   STAT29[4, 7].STAT30 := 0.000000e+000;
   STAT29[4, 7].STAT31 := 0.000000e+000;
   STAT29[4, 7].STAT32 := 0.000000e+000;
   STAT29[4, 8].STAT30 := 0.000000e+000;
   STAT29[4, 8].STAT31 := 0.000000e+000;
   STAT29[4, 8].STAT32 := 0.000000e+000;
   STAT29[4, 9].STAT30 := 0.000000e+000;
   STAT29[4, 9].STAT31 := 0.000000e+000;
   STAT29[4, 9].STAT32 := 0.000000e+000;
   STAT29[4, 10].STAT30 := 0.000000e+000;
   STAT29[4, 10].STAT31 := 0.000000e+000;
   STAT29[4, 10].STAT32 := 0.000000e+000;
   STAT29[5, 1].STAT30 := 0.000000e+000;
   STAT29[5, 1].STAT31 := 0.000000e+000;
   STAT29[5, 1].STAT32 := 0.000000e+000;
   STAT29[5, 2].STAT30 := 0.000000e+000;
   STAT29[5, 2].STAT31 := 0.000000e+000;
   STAT29[5, 2].STAT32 := 0.000000e+000;
   STAT29[5, 3].STAT30 := 0.000000e+000;
   STAT29[5, 3].STAT31 := 0.000000e+000;
   STAT29[5, 3].STAT32 := 0.000000e+000;
   STAT29[5, 4].STAT30 := 0.000000e+000;
   STAT29[5, 4].STAT31 := 0.000000e+000;
   STAT29[5, 4].STAT32 := 0.000000e+000;
   STAT29[5, 5].STAT30 := 0.000000e+000;
   STAT29[5, 5].STAT31 := 0.000000e+000;
   STAT29[5, 5].STAT32 := 0.000000e+000;
   STAT29[5, 6].STAT30 := 0.000000e+000;
   STAT29[5, 6].STAT31 := 0.000000e+000;
   STAT29[5, 6].STAT32 := 0.000000e+000;
   STAT29[5, 7].STAT30 := 0.000000e+000;
   STAT29[5, 7].STAT31 := 0.000000e+000;
   STAT29[5, 7].STAT32 := 0.000000e+000;
   STAT29[5, 8].STAT30 := 0.000000e+000;
   STAT29[5, 8].STAT31 := 0.000000e+000;
   STAT29[5, 8].STAT32 := 0.000000e+000;
   STAT29[5, 9].STAT30 := 0.000000e+000;
   STAT29[5, 9].STAT31 := 0.000000e+000;
   STAT29[5, 9].STAT32 := 0.000000e+000;
   STAT29[5, 10].STAT30 := 0.000000e+000;
   STAT29[5, 10].STAT31 := 0.000000e+000;
   STAT29[5, 10].STAT32 := 0.000000e+000;
   STAT29[6, 1].STAT30 := 0.000000e+000;
   STAT29[6, 1].STAT31 := 0.000000e+000;
   STAT29[6, 1].STAT32 := 0.000000e+000;
   STAT29[6, 2].STAT30 := 0.000000e+000;
   STAT29[6, 2].STAT31 := 0.000000e+000;
   STAT29[6, 2].STAT32 := 0.000000e+000;
   STAT29[6, 3].STAT30 := 0.000000e+000;
   STAT29[6, 3].STAT31 := 0.000000e+000;
   STAT29[6, 3].STAT32 := 0.000000e+000;
   STAT29[6, 4].STAT30 := 0.000000e+000;
   STAT29[6, 4].STAT31 := 0.000000e+000;
   STAT29[6, 4].STAT32 := 0.000000e+000;
   STAT29[6, 5].STAT30 := 0.000000e+000;
   STAT29[6, 5].STAT31 := 0.000000e+000;
   STAT29[6, 5].STAT32 := 0.000000e+000;
   STAT29[6, 6].STAT30 := 0.000000e+000;
   STAT29[6, 6].STAT31 := 0.000000e+000;
   STAT29[6, 6].STAT32 := 0.000000e+000;
   STAT29[6, 7].STAT30 := 0.000000e+000;
   STAT29[6, 7].STAT31 := 0.000000e+000;
   STAT29[6, 7].STAT32 := 0.000000e+000;
   STAT29[6, 8].STAT30 := 0.000000e+000;
   STAT29[6, 8].STAT31 := 0.000000e+000;
   STAT29[6, 8].STAT32 := 0.000000e+000;
   STAT29[6, 9].STAT30 := 0.000000e+000;
   STAT29[6, 9].STAT31 := 0.000000e+000;
   STAT29[6, 9].STAT32 := 0.000000e+000;
   STAT29[6, 10].STAT30 := 0.000000e+000;
   STAT29[6, 10].STAT31 := 0.000000e+000;
   STAT29[6, 10].STAT32 := 0.000000e+000;
   STAT29[7, 1].STAT30 := 0.000000e+000;
   STAT29[7, 1].STAT31 := 0.000000e+000;
   STAT29[7, 1].STAT32 := 0.000000e+000;
   STAT29[7, 2].STAT30 := 0.000000e+000;
   STAT29[7, 2].STAT31 := 0.000000e+000;
   STAT29[7, 2].STAT32 := 0.000000e+000;
   STAT29[7, 3].STAT30 := 0.000000e+000;
   STAT29[7, 3].STAT31 := 0.000000e+000;
   STAT29[7, 3].STAT32 := 0.000000e+000;
   STAT29[7, 4].STAT30 := 0.000000e+000;
   STAT29[7, 4].STAT31 := 0.000000e+000;
   STAT29[7, 4].STAT32 := 0.000000e+000;
   STAT29[7, 5].STAT30 := 0.000000e+000;
   STAT29[7, 5].STAT31 := 0.000000e+000;
   STAT29[7, 5].STAT32 := 0.000000e+000;
   STAT29[7, 6].STAT30 := 0.000000e+000;
   STAT29[7, 6].STAT31 := 0.000000e+000;
   STAT29[7, 6].STAT32 := 0.000000e+000;
   STAT29[7, 7].STAT30 := 0.000000e+000;
   STAT29[7, 7].STAT31 := 0.000000e+000;
   STAT29[7, 7].STAT32 := 0.000000e+000;
   STAT29[7, 8].STAT30 := 0.000000e+000;
   STAT29[7, 8].STAT31 := 0.000000e+000;
   STAT29[7, 8].STAT32 := 0.000000e+000;
   STAT29[7, 9].STAT30 := 0.000000e+000;
   STAT29[7, 9].STAT31 := 0.000000e+000;
   STAT29[7, 9].STAT32 := 0.000000e+000;
   STAT29[7, 10].STAT30 := 0.000000e+000;
   STAT29[7, 10].STAT31 := 0.000000e+000;
   STAT29[7, 10].STAT32 := 0.000000e+000;
   STAT29[8, 1].STAT30 := 0.000000e+000;
   STAT29[8, 1].STAT31 := 0.000000e+000;
   STAT29[8, 1].STAT32 := 0.000000e+000;
   STAT29[8, 2].STAT30 := 0.000000e+000;
   STAT29[8, 2].STAT31 := 0.000000e+000;
   STAT29[8, 2].STAT32 := 0.000000e+000;
   STAT29[8, 3].STAT30 := 0.000000e+000;
   STAT29[8, 3].STAT31 := 0.000000e+000;
   STAT29[8, 3].STAT32 := 0.000000e+000;
   STAT29[8, 4].STAT30 := 0.000000e+000;
   STAT29[8, 4].STAT31 := 0.000000e+000;
   STAT29[8, 4].STAT32 := 0.000000e+000;
   STAT29[8, 5].STAT30 := 0.000000e+000;
   STAT29[8, 5].STAT31 := 0.000000e+000;
   STAT29[8, 5].STAT32 := 0.000000e+000;
   STAT29[8, 6].STAT30 := 0.000000e+000;
   STAT29[8, 6].STAT31 := 0.000000e+000;
   STAT29[8, 6].STAT32 := 0.000000e+000;
   STAT29[8, 7].STAT30 := 0.000000e+000;
   STAT29[8, 7].STAT31 := 0.000000e+000;
   STAT29[8, 7].STAT32 := 0.000000e+000;
   STAT29[8, 8].STAT30 := 0.000000e+000;
   STAT29[8, 8].STAT31 := 0.000000e+000;
   STAT29[8, 8].STAT32 := 0.000000e+000;
   STAT29[8, 9].STAT30 := 0.000000e+000;
   STAT29[8, 9].STAT31 := 0.000000e+000;
   STAT29[8, 9].STAT32 := 0.000000e+000;
   STAT29[8, 10].STAT30 := 0.000000e+000;
   STAT29[8, 10].STAT31 := 0.000000e+000;
   STAT29[8, 10].STAT32 := 0.000000e+000;
   STAT29[9, 1].STAT30 := 0.000000e+000;
   STAT29[9, 1].STAT31 := 0.000000e+000;
   STAT29[9, 1].STAT32 := 0.000000e+000;
   STAT29[9, 2].STAT30 := 0.000000e+000;
   STAT29[9, 2].STAT31 := 0.000000e+000;
   STAT29[9, 2].STAT32 := 0.000000e+000;
   STAT29[9, 3].STAT30 := 0.000000e+000;
   STAT29[9, 3].STAT31 := 0.000000e+000;
   STAT29[9, 3].STAT32 := 0.000000e+000;
   STAT29[9, 4].STAT30 := 0.000000e+000;
   STAT29[9, 4].STAT31 := 0.000000e+000;
   STAT29[9, 4].STAT32 := 0.000000e+000;
   STAT29[9, 5].STAT30 := 0.000000e+000;
   STAT29[9, 5].STAT31 := 0.000000e+000;
   STAT29[9, 5].STAT32 := 0.000000e+000;
   STAT29[9, 6].STAT30 := 0.000000e+000;
   STAT29[9, 6].STAT31 := 0.000000e+000;
   STAT29[9, 6].STAT32 := 0.000000e+000;
   STAT29[9, 7].STAT30 := 0.000000e+000;
   STAT29[9, 7].STAT31 := 0.000000e+000;
   STAT29[9, 7].STAT32 := 0.000000e+000;
   STAT29[9, 8].STAT30 := 0.000000e+000;
   STAT29[9, 8].STAT31 := 0.000000e+000;
   STAT29[9, 8].STAT32 := 0.000000e+000;
   STAT29[9, 9].STAT30 := 0.000000e+000;
   STAT29[9, 9].STAT31 := 0.000000e+000;
   STAT29[9, 9].STAT32 := 0.000000e+000;
   STAT29[9, 10].STAT30 := 0.000000e+000;
   STAT29[9, 10].STAT31 := 0.000000e+000;
   STAT29[9, 10].STAT32 := 0.000000e+000;
   STAT29[10, 1].STAT30 := 0.000000e+000;
   STAT29[10, 1].STAT31 := 0.000000e+000;
   STAT29[10, 1].STAT32 := 0.000000e+000;
   STAT29[10, 2].STAT30 := 0.000000e+000;
   STAT29[10, 2].STAT31 := 0.000000e+000;
   STAT29[10, 2].STAT32 := 0.000000e+000;
   STAT29[10, 3].STAT30 := 0.000000e+000;
   STAT29[10, 3].STAT31 := 0.000000e+000;
   STAT29[10, 3].STAT32 := 0.000000e+000;
   STAT29[10, 4].STAT30 := 0.000000e+000;
   STAT29[10, 4].STAT31 := 0.000000e+000;
   STAT29[10, 4].STAT32 := 0.000000e+000;
   STAT29[10, 5].STAT30 := 0.000000e+000;
   STAT29[10, 5].STAT31 := 0.000000e+000;
   STAT29[10, 5].STAT32 := 0.000000e+000;
   STAT29[10, 6].STAT30 := 0.000000e+000;
   STAT29[10, 6].STAT31 := 0.000000e+000;
   STAT29[10, 6].STAT32 := 0.000000e+000;
   STAT29[10, 7].STAT30 := 0.000000e+000;
   STAT29[10, 7].STAT31 := 0.000000e+000;
   STAT29[10, 7].STAT32 := 0.000000e+000;
   STAT29[10, 8].STAT30 := 0.000000e+000;
   STAT29[10, 8].STAT31 := 0.000000e+000;
   STAT29[10, 8].STAT32 := 0.000000e+000;
   STAT29[10, 9].STAT30 := 0.000000e+000;
   STAT29[10, 9].STAT31 := 0.000000e+000;
   STAT29[10, 9].STAT32 := 0.000000e+000;
   STAT29[10, 10].STAT30 := 0.000000e+000;
   STAT29[10, 10].STAT31 := 0.000000e+000;
   STAT29[10, 10].STAT32 := 0.000000e+000;
   STAT33[1, 1, 1] := 0.000000e+000;
   STAT33[1, 1, 2] := 0.000000e+000;
   STAT33[1, 1, 3] := 0.000000e+000;
   STAT33[1, 1, 4] := 0.000000e+000;
   STAT33[1, 1, 5] := 0.000000e+000;
   STAT33[1, 1, 6] := 0.000000e+000;
   STAT33[1, 1, 7] := 0.000000e+000;
   STAT33[1, 1, 8] := 0.000000e+000;
   STAT33[1, 1, 9] := 0.000000e+000;
   STAT33[1, 1, 10] := 0.000000e+000;
   STAT33[1, 2, 1] := 0.000000e+000;
   STAT33[1, 2, 2] := 0.000000e+000;
   STAT33[1, 2, 3] := 0.000000e+000;
   STAT33[1, 2, 4] := 0.000000e+000;
   STAT33[1, 2, 5] := 0.000000e+000;
   STAT33[1, 2, 6] := 0.000000e+000;
   STAT33[1, 2, 7] := 0.000000e+000;
   STAT33[1, 2, 8] := 0.000000e+000;
   STAT33[1, 2, 9] := 0.000000e+000;
   STAT33[1, 2, 10] := 0.000000e+000;
   STAT33[1, 3, 1] := 0.000000e+000;
   STAT33[1, 3, 2] := 0.000000e+000;
   STAT33[1, 3, 3] := 0.000000e+000;
   STAT33[1, 3, 4] := 0.000000e+000;
   STAT33[1, 3, 5] := 0.000000e+000;
   STAT33[1, 3, 6] := 0.000000e+000;
   STAT33[1, 3, 7] := 0.000000e+000;
   STAT33[1, 3, 8] := 0.000000e+000;
   STAT33[1, 3, 9] := 0.000000e+000;
   STAT33[1, 3, 10] := 0.000000e+000;
   STAT33[1, 4, 1] := 0.000000e+000;
   STAT33[1, 4, 2] := 0.000000e+000;
   STAT33[1, 4, 3] := 0.000000e+000;
   STAT33[1, 4, 4] := 0.000000e+000;
   STAT33[1, 4, 5] := 0.000000e+000;
   STAT33[1, 4, 6] := 0.000000e+000;
   STAT33[1, 4, 7] := 0.000000e+000;
   STAT33[1, 4, 8] := 0.000000e+000;
   STAT33[1, 4, 9] := 0.000000e+000;
   STAT33[1, 4, 10] := 0.000000e+000;
   STAT33[1, 5, 1] := 0.000000e+000;
   STAT33[1, 5, 2] := 0.000000e+000;
   STAT33[1, 5, 3] := 0.000000e+000;
   STAT33[1, 5, 4] := 0.000000e+000;
   STAT33[1, 5, 5] := 0.000000e+000;
   STAT33[1, 5, 6] := 0.000000e+000;
   STAT33[1, 5, 7] := 0.000000e+000;
   STAT33[1, 5, 8] := 0.000000e+000;
   STAT33[1, 5, 9] := 0.000000e+000;
   STAT33[1, 5, 10] := 0.000000e+000;
   STAT33[1, 6, 1] := 0.000000e+000;
   STAT33[1, 6, 2] := 0.000000e+000;
   STAT33[1, 6, 3] := 0.000000e+000;
   STAT33[1, 6, 4] := 0.000000e+000;
   STAT33[1, 6, 5] := 0.000000e+000;
   STAT33[1, 6, 6] := 0.000000e+000;
   STAT33[1, 6, 7] := 0.000000e+000;
   STAT33[1, 6, 8] := 0.000000e+000;
   STAT33[1, 6, 9] := 0.000000e+000;
   STAT33[1, 6, 10] := 0.000000e+000;
   STAT33[1, 7, 1] := 0.000000e+000;
   STAT33[1, 7, 2] := 0.000000e+000;
   STAT33[1, 7, 3] := 0.000000e+000;
   STAT33[1, 7, 4] := 0.000000e+000;
   STAT33[1, 7, 5] := 0.000000e+000;
   STAT33[1, 7, 6] := 0.000000e+000;
   STAT33[1, 7, 7] := 0.000000e+000;
   STAT33[1, 7, 8] := 0.000000e+000;
   STAT33[1, 7, 9] := 0.000000e+000;
   STAT33[1, 7, 10] := 0.000000e+000;
   STAT33[1, 8, 1] := 0.000000e+000;
   STAT33[1, 8, 2] := 0.000000e+000;
   STAT33[1, 8, 3] := 0.000000e+000;
   STAT33[1, 8, 4] := 0.000000e+000;
   STAT33[1, 8, 5] := 0.000000e+000;
   STAT33[1, 8, 6] := 0.000000e+000;
   STAT33[1, 8, 7] := 0.000000e+000;
   STAT33[1, 8, 8] := 0.000000e+000;
   STAT33[1, 8, 9] := 0.000000e+000;
   STAT33[1, 8, 10] := 0.000000e+000;
   STAT33[1, 9, 1] := 0.000000e+000;
   STAT33[1, 9, 2] := 0.000000e+000;
   STAT33[1, 9, 3] := 0.000000e+000;
   STAT33[1, 9, 4] := 0.000000e+000;
   STAT33[1, 9, 5] := 0.000000e+000;
   STAT33[1, 9, 6] := 0.000000e+000;
   STAT33[1, 9, 7] := 0.000000e+000;
   STAT33[1, 9, 8] := 0.000000e+000;
   STAT33[1, 9, 9] := 0.000000e+000;
   STAT33[1, 9, 10] := 0.000000e+000;
   STAT33[1, 10, 1] := 0.000000e+000;
   STAT33[1, 10, 2] := 0.000000e+000;
   STAT33[1, 10, 3] := 0.000000e+000;
   STAT33[1, 10, 4] := 0.000000e+000;
   STAT33[1, 10, 5] := 0.000000e+000;
   STAT33[1, 10, 6] := 0.000000e+000;
   STAT33[1, 10, 7] := 0.000000e+000;
   STAT33[1, 10, 8] := 0.000000e+000;
   STAT33[1, 10, 9] := 0.000000e+000;
   STAT33[1, 10, 10] := 0.000000e+000;
   STAT33[2, 1, 1] := 0.000000e+000;
   STAT33[2, 1, 2] := 0.000000e+000;
   STAT33[2, 1, 3] := 0.000000e+000;
   STAT33[2, 1, 4] := 0.000000e+000;
   STAT33[2, 1, 5] := 0.000000e+000;
   STAT33[2, 1, 6] := 0.000000e+000;
   STAT33[2, 1, 7] := 0.000000e+000;
   STAT33[2, 1, 8] := 0.000000e+000;
   STAT33[2, 1, 9] := 0.000000e+000;
   STAT33[2, 1, 10] := 0.000000e+000;
   STAT33[2, 2, 1] := 0.000000e+000;
   STAT33[2, 2, 2] := 0.000000e+000;
   STAT33[2, 2, 3] := 0.000000e+000;
   STAT33[2, 2, 4] := 0.000000e+000;
   STAT33[2, 2, 5] := 0.000000e+000;
   STAT33[2, 2, 6] := 0.000000e+000;
   STAT33[2, 2, 7] := 0.000000e+000;
   STAT33[2, 2, 8] := 0.000000e+000;
   STAT33[2, 2, 9] := 0.000000e+000;
   STAT33[2, 2, 10] := 0.000000e+000;
   STAT33[2, 3, 1] := 0.000000e+000;
   STAT33[2, 3, 2] := 0.000000e+000;
   STAT33[2, 3, 3] := 0.000000e+000;
   STAT33[2, 3, 4] := 0.000000e+000;
   STAT33[2, 3, 5] := 0.000000e+000;
   STAT33[2, 3, 6] := 0.000000e+000;
   STAT33[2, 3, 7] := 0.000000e+000;
   STAT33[2, 3, 8] := 0.000000e+000;
   STAT33[2, 3, 9] := 0.000000e+000;
   STAT33[2, 3, 10] := 0.000000e+000;
   STAT33[2, 4, 1] := 0.000000e+000;
   STAT33[2, 4, 2] := 0.000000e+000;
   STAT33[2, 4, 3] := 0.000000e+000;
   STAT33[2, 4, 4] := 0.000000e+000;
   STAT33[2, 4, 5] := 0.000000e+000;
   STAT33[2, 4, 6] := 0.000000e+000;
   STAT33[2, 4, 7] := 0.000000e+000;
   STAT33[2, 4, 8] := 0.000000e+000;
   STAT33[2, 4, 9] := 0.000000e+000;
   STAT33[2, 4, 10] := 0.000000e+000;
   STAT33[2, 5, 1] := 0.000000e+000;
   STAT33[2, 5, 2] := 0.000000e+000;
   STAT33[2, 5, 3] := 0.000000e+000;
   STAT33[2, 5, 4] := 0.000000e+000;
   STAT33[2, 5, 5] := 0.000000e+000;
   STAT33[2, 5, 6] := 0.000000e+000;
   STAT33[2, 5, 7] := 0.000000e+000;
   STAT33[2, 5, 8] := 0.000000e+000;
   STAT33[2, 5, 9] := 0.000000e+000;
   STAT33[2, 5, 10] := 0.000000e+000;
   STAT33[2, 6, 1] := 0.000000e+000;
   STAT33[2, 6, 2] := 0.000000e+000;
   STAT33[2, 6, 3] := 0.000000e+000;
   STAT33[2, 6, 4] := 0.000000e+000;
   STAT33[2, 6, 5] := 0.000000e+000;
   STAT33[2, 6, 6] := 0.000000e+000;
   STAT33[2, 6, 7] := 0.000000e+000;
   STAT33[2, 6, 8] := 0.000000e+000;
   STAT33[2, 6, 9] := 0.000000e+000;
   STAT33[2, 6, 10] := 0.000000e+000;
   STAT33[2, 7, 1] := 0.000000e+000;
   STAT33[2, 7, 2] := 0.000000e+000;
   STAT33[2, 7, 3] := 0.000000e+000;
   STAT33[2, 7, 4] := 0.000000e+000;
   STAT33[2, 7, 5] := 0.000000e+000;
   STAT33[2, 7, 6] := 0.000000e+000;
   STAT33[2, 7, 7] := 0.000000e+000;
   STAT33[2, 7, 8] := 0.000000e+000;
   STAT33[2, 7, 9] := 0.000000e+000;
   STAT33[2, 7, 10] := 0.000000e+000;
   STAT33[2, 8, 1] := 0.000000e+000;
   STAT33[2, 8, 2] := 0.000000e+000;
   STAT33[2, 8, 3] := 0.000000e+000;
   STAT33[2, 8, 4] := 0.000000e+000;
   STAT33[2, 8, 5] := 0.000000e+000;
   STAT33[2, 8, 6] := 0.000000e+000;
   STAT33[2, 8, 7] := 0.000000e+000;
   STAT33[2, 8, 8] := 0.000000e+000;
   STAT33[2, 8, 9] := 0.000000e+000;
   STAT33[2, 8, 10] := 0.000000e+000;
   STAT33[2, 9, 1] := 0.000000e+000;
   STAT33[2, 9, 2] := 0.000000e+000;
   STAT33[2, 9, 3] := 0.000000e+000;
   STAT33[2, 9, 4] := 0.000000e+000;
   STAT33[2, 9, 5] := 0.000000e+000;
   STAT33[2, 9, 6] := 0.000000e+000;
   STAT33[2, 9, 7] := 0.000000e+000;
   STAT33[2, 9, 8] := 0.000000e+000;
   STAT33[2, 9, 9] := 0.000000e+000;
   STAT33[2, 9, 10] := 0.000000e+000;
   STAT33[2, 10, 1] := 0.000000e+000;
   STAT33[2, 10, 2] := 0.000000e+000;
   STAT33[2, 10, 3] := 0.000000e+000;
   STAT33[2, 10, 4] := 0.000000e+000;
   STAT33[2, 10, 5] := 0.000000e+000;
   STAT33[2, 10, 6] := 0.000000e+000;
   STAT33[2, 10, 7] := 0.000000e+000;
   STAT33[2, 10, 8] := 0.000000e+000;
   STAT33[2, 10, 9] := 0.000000e+000;
   STAT33[2, 10, 10] := 0.000000e+000;
   STAT33[3, 1, 1] := 0.000000e+000;
   STAT33[3, 1, 2] := 0.000000e+000;
   STAT33[3, 1, 3] := 0.000000e+000;
   STAT33[3, 1, 4] := 0.000000e+000;
   STAT33[3, 1, 5] := 0.000000e+000;
   STAT33[3, 1, 6] := 0.000000e+000;
   STAT33[3, 1, 7] := 0.000000e+000;
   STAT33[3, 1, 8] := 0.000000e+000;
   STAT33[3, 1, 9] := 0.000000e+000;
   STAT33[3, 1, 10] := 0.000000e+000;
   STAT33[3, 2, 1] := 0.000000e+000;
   STAT33[3, 2, 2] := 0.000000e+000;
   STAT33[3, 2, 3] := 0.000000e+000;
   STAT33[3, 2, 4] := 0.000000e+000;
   STAT33[3, 2, 5] := 0.000000e+000;
   STAT33[3, 2, 6] := 0.000000e+000;
   STAT33[3, 2, 7] := 0.000000e+000;
   STAT33[3, 2, 8] := 0.000000e+000;
   STAT33[3, 2, 9] := 0.000000e+000;
   STAT33[3, 2, 10] := 0.000000e+000;
   STAT33[3, 3, 1] := 0.000000e+000;
   STAT33[3, 3, 2] := 0.000000e+000;
   STAT33[3, 3, 3] := 0.000000e+000;
   STAT33[3, 3, 4] := 0.000000e+000;
   STAT33[3, 3, 5] := 0.000000e+000;
   STAT33[3, 3, 6] := 0.000000e+000;
   STAT33[3, 3, 7] := 0.000000e+000;
   STAT33[3, 3, 8] := 0.000000e+000;
   STAT33[3, 3, 9] := 0.000000e+000;
   STAT33[3, 3, 10] := 0.000000e+000;
   STAT33[3, 4, 1] := 0.000000e+000;
   STAT33[3, 4, 2] := 0.000000e+000;
   STAT33[3, 4, 3] := 0.000000e+000;
   STAT33[3, 4, 4] := 0.000000e+000;
   STAT33[3, 4, 5] := 0.000000e+000;
   STAT33[3, 4, 6] := 0.000000e+000;
   STAT33[3, 4, 7] := 0.000000e+000;
   STAT33[3, 4, 8] := 0.000000e+000;
   STAT33[3, 4, 9] := 0.000000e+000;
   STAT33[3, 4, 10] := 0.000000e+000;
   STAT33[3, 5, 1] := 0.000000e+000;
   STAT33[3, 5, 2] := 0.000000e+000;
   STAT33[3, 5, 3] := 0.000000e+000;
   STAT33[3, 5, 4] := 0.000000e+000;
   STAT33[3, 5, 5] := 0.000000e+000;
   STAT33[3, 5, 6] := 0.000000e+000;
   STAT33[3, 5, 7] := 0.000000e+000;
   STAT33[3, 5, 8] := 0.000000e+000;
   STAT33[3, 5, 9] := 0.000000e+000;
   STAT33[3, 5, 10] := 0.000000e+000;
   STAT33[3, 6, 1] := 0.000000e+000;
   STAT33[3, 6, 2] := 0.000000e+000;
   STAT33[3, 6, 3] := 0.000000e+000;
   STAT33[3, 6, 4] := 0.000000e+000;
   STAT33[3, 6, 5] := 0.000000e+000;
   STAT33[3, 6, 6] := 0.000000e+000;
   STAT33[3, 6, 7] := 0.000000e+000;
   STAT33[3, 6, 8] := 0.000000e+000;
   STAT33[3, 6, 9] := 0.000000e+000;
   STAT33[3, 6, 10] := 0.000000e+000;
   STAT33[3, 7, 1] := 0.000000e+000;
   STAT33[3, 7, 2] := 0.000000e+000;
   STAT33[3, 7, 3] := 0.000000e+000;
   STAT33[3, 7, 4] := 0.000000e+000;
   STAT33[3, 7, 5] := 0.000000e+000;
   STAT33[3, 7, 6] := 0.000000e+000;
   STAT33[3, 7, 7] := 0.000000e+000;
   STAT33[3, 7, 8] := 0.000000e+000;
   STAT33[3, 7, 9] := 0.000000e+000;
   STAT33[3, 7, 10] := 0.000000e+000;
   STAT33[3, 8, 1] := 0.000000e+000;
   STAT33[3, 8, 2] := 0.000000e+000;
   STAT33[3, 8, 3] := 0.000000e+000;
   STAT33[3, 8, 4] := 0.000000e+000;
   STAT33[3, 8, 5] := 0.000000e+000;
   STAT33[3, 8, 6] := 0.000000e+000;
   STAT33[3, 8, 7] := 0.000000e+000;
   STAT33[3, 8, 8] := 0.000000e+000;
   STAT33[3, 8, 9] := 0.000000e+000;
   STAT33[3, 8, 10] := 0.000000e+000;
   STAT33[3, 9, 1] := 0.000000e+000;
   STAT33[3, 9, 2] := 0.000000e+000;
   STAT33[3, 9, 3] := 0.000000e+000;
   STAT33[3, 9, 4] := 0.000000e+000;
   STAT33[3, 9, 5] := 0.000000e+000;
   STAT33[3, 9, 6] := 0.000000e+000;
   STAT33[3, 9, 7] := 0.000000e+000;
   STAT33[3, 9, 8] := 0.000000e+000;
   STAT33[3, 9, 9] := 0.000000e+000;
   STAT33[3, 9, 10] := 0.000000e+000;
   STAT33[3, 10, 1] := 0.000000e+000;
   STAT33[3, 10, 2] := 0.000000e+000;
   STAT33[3, 10, 3] := 0.000000e+000;
   STAT33[3, 10, 4] := 0.000000e+000;
   STAT33[3, 10, 5] := 0.000000e+000;
   STAT33[3, 10, 6] := 0.000000e+000;
   STAT33[3, 10, 7] := 0.000000e+000;
   STAT33[3, 10, 8] := 0.000000e+000;
   STAT33[3, 10, 9] := 0.000000e+000;
   STAT33[3, 10, 10] := 0.000000e+000;
   STAT33[4, 1, 1] := 0.000000e+000;
   STAT33[4, 1, 2] := 0.000000e+000;
   STAT33[4, 1, 3] := 0.000000e+000;
   STAT33[4, 1, 4] := 0.000000e+000;
   STAT33[4, 1, 5] := 0.000000e+000;
   STAT33[4, 1, 6] := 0.000000e+000;
   STAT33[4, 1, 7] := 0.000000e+000;
   STAT33[4, 1, 8] := 0.000000e+000;
   STAT33[4, 1, 9] := 0.000000e+000;
   STAT33[4, 1, 10] := 0.000000e+000;
   STAT33[4, 2, 1] := 0.000000e+000;
   STAT33[4, 2, 2] := 0.000000e+000;
   STAT33[4, 2, 3] := 0.000000e+000;
   STAT33[4, 2, 4] := 0.000000e+000;
   STAT33[4, 2, 5] := 0.000000e+000;
   STAT33[4, 2, 6] := 0.000000e+000;
   STAT33[4, 2, 7] := 0.000000e+000;
   STAT33[4, 2, 8] := 0.000000e+000;
   STAT33[4, 2, 9] := 0.000000e+000;
   STAT33[4, 2, 10] := 0.000000e+000;
   STAT33[4, 3, 1] := 0.000000e+000;
   STAT33[4, 3, 2] := 0.000000e+000;
   STAT33[4, 3, 3] := 0.000000e+000;
   STAT33[4, 3, 4] := 0.000000e+000;
   STAT33[4, 3, 5] := 0.000000e+000;
   STAT33[4, 3, 6] := 0.000000e+000;
   STAT33[4, 3, 7] := 0.000000e+000;
   STAT33[4, 3, 8] := 0.000000e+000;
   STAT33[4, 3, 9] := 0.000000e+000;
   STAT33[4, 3, 10] := 0.000000e+000;
   STAT33[4, 4, 1] := 0.000000e+000;
   STAT33[4, 4, 2] := 0.000000e+000;
   STAT33[4, 4, 3] := 0.000000e+000;
   STAT33[4, 4, 4] := 0.000000e+000;
   STAT33[4, 4, 5] := 0.000000e+000;
   STAT33[4, 4, 6] := 0.000000e+000;
   STAT33[4, 4, 7] := 0.000000e+000;
   STAT33[4, 4, 8] := 0.000000e+000;
   STAT33[4, 4, 9] := 0.000000e+000;
   STAT33[4, 4, 10] := 0.000000e+000;
   STAT33[4, 5, 1] := 0.000000e+000;
   STAT33[4, 5, 2] := 0.000000e+000;
   STAT33[4, 5, 3] := 0.000000e+000;
   STAT33[4, 5, 4] := 0.000000e+000;
   STAT33[4, 5, 5] := 0.000000e+000;
   STAT33[4, 5, 6] := 0.000000e+000;
   STAT33[4, 5, 7] := 0.000000e+000;
   STAT33[4, 5, 8] := 0.000000e+000;
   STAT33[4, 5, 9] := 0.000000e+000;
   STAT33[4, 5, 10] := 0.000000e+000;
   STAT33[4, 6, 1] := 0.000000e+000;
   STAT33[4, 6, 2] := 0.000000e+000;
   STAT33[4, 6, 3] := 0.000000e+000;
   STAT33[4, 6, 4] := 0.000000e+000;
   STAT33[4, 6, 5] := 0.000000e+000;
   STAT33[4, 6, 6] := 0.000000e+000;
   STAT33[4, 6, 7] := 0.000000e+000;
   STAT33[4, 6, 8] := 0.000000e+000;
   STAT33[4, 6, 9] := 0.000000e+000;
   STAT33[4, 6, 10] := 0.000000e+000;
   STAT33[4, 7, 1] := 0.000000e+000;
   STAT33[4, 7, 2] := 0.000000e+000;
   STAT33[4, 7, 3] := 0.000000e+000;
   STAT33[4, 7, 4] := 0.000000e+000;
   STAT33[4, 7, 5] := 0.000000e+000;
   STAT33[4, 7, 6] := 0.000000e+000;
   STAT33[4, 7, 7] := 0.000000e+000;
   STAT33[4, 7, 8] := 0.000000e+000;
   STAT33[4, 7, 9] := 0.000000e+000;
   STAT33[4, 7, 10] := 0.000000e+000;
   STAT33[4, 8, 1] := 0.000000e+000;
   STAT33[4, 8, 2] := 0.000000e+000;
   STAT33[4, 8, 3] := 0.000000e+000;
   STAT33[4, 8, 4] := 0.000000e+000;
   STAT33[4, 8, 5] := 0.000000e+000;
   STAT33[4, 8, 6] := 0.000000e+000;
   STAT33[4, 8, 7] := 0.000000e+000;
   STAT33[4, 8, 8] := 0.000000e+000;
   STAT33[4, 8, 9] := 0.000000e+000;
   STAT33[4, 8, 10] := 0.000000e+000;
   STAT33[4, 9, 1] := 0.000000e+000;
   STAT33[4, 9, 2] := 0.000000e+000;
   STAT33[4, 9, 3] := 0.000000e+000;
   STAT33[4, 9, 4] := 0.000000e+000;
   STAT33[4, 9, 5] := 0.000000e+000;
   STAT33[4, 9, 6] := 0.000000e+000;
   STAT33[4, 9, 7] := 0.000000e+000;
   STAT33[4, 9, 8] := 0.000000e+000;
   STAT33[4, 9, 9] := 0.000000e+000;
   STAT33[4, 9, 10] := 0.000000e+000;
   STAT33[4, 10, 1] := 0.000000e+000;
   STAT33[4, 10, 2] := 0.000000e+000;
   STAT33[4, 10, 3] := 0.000000e+000;
   STAT33[4, 10, 4] := 0.000000e+000;
   STAT33[4, 10, 5] := 0.000000e+000;
   STAT33[4, 10, 6] := 0.000000e+000;
   STAT33[4, 10, 7] := 0.000000e+000;
   STAT33[4, 10, 8] := 0.000000e+000;
   STAT33[4, 10, 9] := 0.000000e+000;
   STAT33[4, 10, 10] := 0.000000e+000;
   STAT33[5, 1, 1] := 0.000000e+000;
   STAT33[5, 1, 2] := 0.000000e+000;
   STAT33[5, 1, 3] := 0.000000e+000;
   STAT33[5, 1, 4] := 0.000000e+000;
   STAT33[5, 1, 5] := 0.000000e+000;
   STAT33[5, 1, 6] := 0.000000e+000;
   STAT33[5, 1, 7] := 0.000000e+000;
   STAT33[5, 1, 8] := 0.000000e+000;
   STAT33[5, 1, 9] := 0.000000e+000;
   STAT33[5, 1, 10] := 0.000000e+000;
   STAT33[5, 2, 1] := 0.000000e+000;
   STAT33[5, 2, 2] := 0.000000e+000;
   STAT33[5, 2, 3] := 0.000000e+000;
   STAT33[5, 2, 4] := 0.000000e+000;
   STAT33[5, 2, 5] := 0.000000e+000;
   STAT33[5, 2, 6] := 0.000000e+000;
   STAT33[5, 2, 7] := 0.000000e+000;
   STAT33[5, 2, 8] := 0.000000e+000;
   STAT33[5, 2, 9] := 0.000000e+000;
   STAT33[5, 2, 10] := 0.000000e+000;
   STAT33[5, 3, 1] := 0.000000e+000;
   STAT33[5, 3, 2] := 0.000000e+000;
   STAT33[5, 3, 3] := 0.000000e+000;
   STAT33[5, 3, 4] := 0.000000e+000;
   STAT33[5, 3, 5] := 0.000000e+000;
   STAT33[5, 3, 6] := 0.000000e+000;
   STAT33[5, 3, 7] := 0.000000e+000;
   STAT33[5, 3, 8] := 0.000000e+000;
   STAT33[5, 3, 9] := 0.000000e+000;
   STAT33[5, 3, 10] := 0.000000e+000;
   STAT33[5, 4, 1] := 0.000000e+000;
   STAT33[5, 4, 2] := 0.000000e+000;
   STAT33[5, 4, 3] := 0.000000e+000;
   STAT33[5, 4, 4] := 0.000000e+000;
   STAT33[5, 4, 5] := 0.000000e+000;
   STAT33[5, 4, 6] := 0.000000e+000;
   STAT33[5, 4, 7] := 0.000000e+000;
   STAT33[5, 4, 8] := 0.000000e+000;
   STAT33[5, 4, 9] := 0.000000e+000;
   STAT33[5, 4, 10] := 0.000000e+000;
   STAT33[5, 5, 1] := 0.000000e+000;
   STAT33[5, 5, 2] := 0.000000e+000;
   STAT33[5, 5, 3] := 0.000000e+000;
   STAT33[5, 5, 4] := 0.000000e+000;
   STAT33[5, 5, 5] := 0.000000e+000;
   STAT33[5, 5, 6] := 0.000000e+000;
   STAT33[5, 5, 7] := 0.000000e+000;
   STAT33[5, 5, 8] := 0.000000e+000;
   STAT33[5, 5, 9] := 0.000000e+000;
   STAT33[5, 5, 10] := 0.000000e+000;
   STAT33[5, 6, 1] := 0.000000e+000;
   STAT33[5, 6, 2] := 0.000000e+000;
   STAT33[5, 6, 3] := 0.000000e+000;
   STAT33[5, 6, 4] := 0.000000e+000;
   STAT33[5, 6, 5] := 0.000000e+000;
   STAT33[5, 6, 6] := 0.000000e+000;
   STAT33[5, 6, 7] := 0.000000e+000;
   STAT33[5, 6, 8] := 0.000000e+000;
   STAT33[5, 6, 9] := 0.000000e+000;
   STAT33[5, 6, 10] := 0.000000e+000;
   STAT33[5, 7, 1] := 0.000000e+000;
   STAT33[5, 7, 2] := 0.000000e+000;
   STAT33[5, 7, 3] := 0.000000e+000;
   STAT33[5, 7, 4] := 0.000000e+000;
   STAT33[5, 7, 5] := 0.000000e+000;
   STAT33[5, 7, 6] := 0.000000e+000;
   STAT33[5, 7, 7] := 0.000000e+000;
   STAT33[5, 7, 8] := 0.000000e+000;
   STAT33[5, 7, 9] := 0.000000e+000;
   STAT33[5, 7, 10] := 0.000000e+000;
   STAT33[5, 8, 1] := 0.000000e+000;
   STAT33[5, 8, 2] := 0.000000e+000;
   STAT33[5, 8, 3] := 0.000000e+000;
   STAT33[5, 8, 4] := 0.000000e+000;
   STAT33[5, 8, 5] := 0.000000e+000;
   STAT33[5, 8, 6] := 0.000000e+000;
   STAT33[5, 8, 7] := 0.000000e+000;
   STAT33[5, 8, 8] := 0.000000e+000;
   STAT33[5, 8, 9] := 0.000000e+000;
   STAT33[5, 8, 10] := 0.000000e+000;
   STAT33[5, 9, 1] := 0.000000e+000;
   STAT33[5, 9, 2] := 0.000000e+000;
   STAT33[5, 9, 3] := 0.000000e+000;
   STAT33[5, 9, 4] := 0.000000e+000;
   STAT33[5, 9, 5] := 0.000000e+000;
   STAT33[5, 9, 6] := 0.000000e+000;
   STAT33[5, 9, 7] := 0.000000e+000;
   STAT33[5, 9, 8] := 0.000000e+000;
   STAT33[5, 9, 9] := 0.000000e+000;
   STAT33[5, 9, 10] := 0.000000e+000;
   STAT33[5, 10, 1] := 0.000000e+000;
   STAT33[5, 10, 2] := 0.000000e+000;
   STAT33[5, 10, 3] := 0.000000e+000;
   STAT33[5, 10, 4] := 0.000000e+000;
   STAT33[5, 10, 5] := 0.000000e+000;
   STAT33[5, 10, 6] := 0.000000e+000;
   STAT33[5, 10, 7] := 0.000000e+000;
   STAT33[5, 10, 8] := 0.000000e+000;
   STAT33[5, 10, 9] := 0.000000e+000;
   STAT33[5, 10, 10] := 0.000000e+000;
   STAT33[6, 1, 1] := 0.000000e+000;
   STAT33[6, 1, 2] := 0.000000e+000;
   STAT33[6, 1, 3] := 0.000000e+000;
   STAT33[6, 1, 4] := 0.000000e+000;
   STAT33[6, 1, 5] := 0.000000e+000;
   STAT33[6, 1, 6] := 0.000000e+000;
   STAT33[6, 1, 7] := 0.000000e+000;
   STAT33[6, 1, 8] := 0.000000e+000;
   STAT33[6, 1, 9] := 0.000000e+000;
   STAT33[6, 1, 10] := 0.000000e+000;
   STAT33[6, 2, 1] := 0.000000e+000;
   STAT33[6, 2, 2] := 0.000000e+000;
   STAT33[6, 2, 3] := 0.000000e+000;
   STAT33[6, 2, 4] := 0.000000e+000;
   STAT33[6, 2, 5] := 0.000000e+000;
   STAT33[6, 2, 6] := 0.000000e+000;
   STAT33[6, 2, 7] := 0.000000e+000;
   STAT33[6, 2, 8] := 0.000000e+000;
   STAT33[6, 2, 9] := 0.000000e+000;
   STAT33[6, 2, 10] := 0.000000e+000;
   STAT33[6, 3, 1] := 0.000000e+000;
   STAT33[6, 3, 2] := 0.000000e+000;
   STAT33[6, 3, 3] := 0.000000e+000;
   STAT33[6, 3, 4] := 0.000000e+000;
   STAT33[6, 3, 5] := 0.000000e+000;
   STAT33[6, 3, 6] := 0.000000e+000;
   STAT33[6, 3, 7] := 0.000000e+000;
   STAT33[6, 3, 8] := 0.000000e+000;
   STAT33[6, 3, 9] := 0.000000e+000;
   STAT33[6, 3, 10] := 0.000000e+000;
   STAT33[6, 4, 1] := 0.000000e+000;
   STAT33[6, 4, 2] := 0.000000e+000;
   STAT33[6, 4, 3] := 0.000000e+000;
   STAT33[6, 4, 4] := 0.000000e+000;
   STAT33[6, 4, 5] := 0.000000e+000;
   STAT33[6, 4, 6] := 0.000000e+000;
   STAT33[6, 4, 7] := 0.000000e+000;
   STAT33[6, 4, 8] := 0.000000e+000;
   STAT33[6, 4, 9] := 0.000000e+000;
   STAT33[6, 4, 10] := 0.000000e+000;
   STAT33[6, 5, 1] := 0.000000e+000;
   STAT33[6, 5, 2] := 0.000000e+000;
   STAT33[6, 5, 3] := 0.000000e+000;
   STAT33[6, 5, 4] := 0.000000e+000;
   STAT33[6, 5, 5] := 0.000000e+000;
   STAT33[6, 5, 6] := 0.000000e+000;
   STAT33[6, 5, 7] := 0.000000e+000;
   STAT33[6, 5, 8] := 0.000000e+000;
   STAT33[6, 5, 9] := 0.000000e+000;
   STAT33[6, 5, 10] := 0.000000e+000;
   STAT33[6, 6, 1] := 0.000000e+000;
   STAT33[6, 6, 2] := 0.000000e+000;
   STAT33[6, 6, 3] := 0.000000e+000;
   STAT33[6, 6, 4] := 0.000000e+000;
   STAT33[6, 6, 5] := 0.000000e+000;
   STAT33[6, 6, 6] := 0.000000e+000;
   STAT33[6, 6, 7] := 0.000000e+000;
   STAT33[6, 6, 8] := 0.000000e+000;
   STAT33[6, 6, 9] := 0.000000e+000;
   STAT33[6, 6, 10] := 0.000000e+000;
   STAT33[6, 7, 1] := 0.000000e+000;
   STAT33[6, 7, 2] := 0.000000e+000;
   STAT33[6, 7, 3] := 0.000000e+000;
   STAT33[6, 7, 4] := 0.000000e+000;
   STAT33[6, 7, 5] := 0.000000e+000;
   STAT33[6, 7, 6] := 0.000000e+000;
   STAT33[6, 7, 7] := 0.000000e+000;
   STAT33[6, 7, 8] := 0.000000e+000;
   STAT33[6, 7, 9] := 0.000000e+000;
   STAT33[6, 7, 10] := 0.000000e+000;
   STAT33[6, 8, 1] := 0.000000e+000;
   STAT33[6, 8, 2] := 0.000000e+000;
   STAT33[6, 8, 3] := 0.000000e+000;
   STAT33[6, 8, 4] := 0.000000e+000;
   STAT33[6, 8, 5] := 0.000000e+000;
   STAT33[6, 8, 6] := 0.000000e+000;
   STAT33[6, 8, 7] := 0.000000e+000;
   STAT33[6, 8, 8] := 0.000000e+000;
   STAT33[6, 8, 9] := 0.000000e+000;
   STAT33[6, 8, 10] := 0.000000e+000;
   STAT33[6, 9, 1] := 0.000000e+000;
   STAT33[6, 9, 2] := 0.000000e+000;
   STAT33[6, 9, 3] := 0.000000e+000;
   STAT33[6, 9, 4] := 0.000000e+000;
   STAT33[6, 9, 5] := 0.000000e+000;
   STAT33[6, 9, 6] := 0.000000e+000;
   STAT33[6, 9, 7] := 0.000000e+000;
   STAT33[6, 9, 8] := 0.000000e+000;
   STAT33[6, 9, 9] := 0.000000e+000;
   STAT33[6, 9, 10] := 0.000000e+000;
   STAT33[6, 10, 1] := 0.000000e+000;
   STAT33[6, 10, 2] := 0.000000e+000;
   STAT33[6, 10, 3] := 0.000000e+000;
   STAT33[6, 10, 4] := 0.000000e+000;
   STAT33[6, 10, 5] := 0.000000e+000;
   STAT33[6, 10, 6] := 0.000000e+000;
   STAT33[6, 10, 7] := 0.000000e+000;
   STAT33[6, 10, 8] := 0.000000e+000;
   STAT33[6, 10, 9] := 0.000000e+000;
   STAT33[6, 10, 10] := 0.000000e+000;
   STAT33[7, 1, 1] := 0.000000e+000;
   STAT33[7, 1, 2] := 0.000000e+000;
   STAT33[7, 1, 3] := 0.000000e+000;
   STAT33[7, 1, 4] := 0.000000e+000;
   STAT33[7, 1, 5] := 0.000000e+000;
   STAT33[7, 1, 6] := 0.000000e+000;
   STAT33[7, 1, 7] := 0.000000e+000;
   STAT33[7, 1, 8] := 0.000000e+000;
   STAT33[7, 1, 9] := 0.000000e+000;
   STAT33[7, 1, 10] := 0.000000e+000;
   STAT33[7, 2, 1] := 0.000000e+000;
   STAT33[7, 2, 2] := 0.000000e+000;
   STAT33[7, 2, 3] := 0.000000e+000;
   STAT33[7, 2, 4] := 0.000000e+000;
   STAT33[7, 2, 5] := 0.000000e+000;
   STAT33[7, 2, 6] := 0.000000e+000;
   STAT33[7, 2, 7] := 0.000000e+000;
   STAT33[7, 2, 8] := 0.000000e+000;
   STAT33[7, 2, 9] := 0.000000e+000;
   STAT33[7, 2, 10] := 0.000000e+000;
   STAT33[7, 3, 1] := 0.000000e+000;
   STAT33[7, 3, 2] := 0.000000e+000;
   STAT33[7, 3, 3] := 0.000000e+000;
   STAT33[7, 3, 4] := 0.000000e+000;
   STAT33[7, 3, 5] := 0.000000e+000;
   STAT33[7, 3, 6] := 0.000000e+000;
   STAT33[7, 3, 7] := 0.000000e+000;
   STAT33[7, 3, 8] := 0.000000e+000;
   STAT33[7, 3, 9] := 0.000000e+000;
   STAT33[7, 3, 10] := 0.000000e+000;
   STAT33[7, 4, 1] := 0.000000e+000;
   STAT33[7, 4, 2] := 0.000000e+000;
   STAT33[7, 4, 3] := 0.000000e+000;
   STAT33[7, 4, 4] := 0.000000e+000;
   STAT33[7, 4, 5] := 0.000000e+000;
   STAT33[7, 4, 6] := 0.000000e+000;
   STAT33[7, 4, 7] := 0.000000e+000;
   STAT33[7, 4, 8] := 0.000000e+000;
   STAT33[7, 4, 9] := 0.000000e+000;
   STAT33[7, 4, 10] := 0.000000e+000;
   STAT33[7, 5, 1] := 0.000000e+000;
   STAT33[7, 5, 2] := 0.000000e+000;
   STAT33[7, 5, 3] := 0.000000e+000;
   STAT33[7, 5, 4] := 0.000000e+000;
   STAT33[7, 5, 5] := 0.000000e+000;
   STAT33[7, 5, 6] := 0.000000e+000;
   STAT33[7, 5, 7] := 0.000000e+000;
   STAT33[7, 5, 8] := 0.000000e+000;
   STAT33[7, 5, 9] := 0.000000e+000;
   STAT33[7, 5, 10] := 0.000000e+000;
   STAT33[7, 6, 1] := 0.000000e+000;
   STAT33[7, 6, 2] := 0.000000e+000;
   STAT33[7, 6, 3] := 0.000000e+000;
   STAT33[7, 6, 4] := 0.000000e+000;
   STAT33[7, 6, 5] := 0.000000e+000;
   STAT33[7, 6, 6] := 0.000000e+000;
   STAT33[7, 6, 7] := 0.000000e+000;
   STAT33[7, 6, 8] := 0.000000e+000;
   STAT33[7, 6, 9] := 0.000000e+000;
   STAT33[7, 6, 10] := 0.000000e+000;
   STAT33[7, 7, 1] := 0.000000e+000;
   STAT33[7, 7, 2] := 0.000000e+000;
   STAT33[7, 7, 3] := 0.000000e+000;
   STAT33[7, 7, 4] := 0.000000e+000;
   STAT33[7, 7, 5] := 0.000000e+000;
   STAT33[7, 7, 6] := 0.000000e+000;
   STAT33[7, 7, 7] := 0.000000e+000;
   STAT33[7, 7, 8] := 0.000000e+000;
   STAT33[7, 7, 9] := 0.000000e+000;
   STAT33[7, 7, 10] := 0.000000e+000;
   STAT33[7, 8, 1] := 0.000000e+000;
   STAT33[7, 8, 2] := 0.000000e+000;
   STAT33[7, 8, 3] := 0.000000e+000;
   STAT33[7, 8, 4] := 0.000000e+000;
   STAT33[7, 8, 5] := 0.000000e+000;
   STAT33[7, 8, 6] := 0.000000e+000;
   STAT33[7, 8, 7] := 0.000000e+000;
   STAT33[7, 8, 8] := 0.000000e+000;
   STAT33[7, 8, 9] := 0.000000e+000;
   STAT33[7, 8, 10] := 0.000000e+000;
   STAT33[7, 9, 1] := 0.000000e+000;
   STAT33[7, 9, 2] := 0.000000e+000;
   STAT33[7, 9, 3] := 0.000000e+000;
   STAT33[7, 9, 4] := 0.000000e+000;
   STAT33[7, 9, 5] := 0.000000e+000;
   STAT33[7, 9, 6] := 0.000000e+000;
   STAT33[7, 9, 7] := 0.000000e+000;
   STAT33[7, 9, 8] := 0.000000e+000;
   STAT33[7, 9, 9] := 0.000000e+000;
   STAT33[7, 9, 10] := 0.000000e+000;
   STAT33[7, 10, 1] := 0.000000e+000;
   STAT33[7, 10, 2] := 0.000000e+000;
   STAT33[7, 10, 3] := 0.000000e+000;
   STAT33[7, 10, 4] := 0.000000e+000;
   STAT33[7, 10, 5] := 0.000000e+000;
   STAT33[7, 10, 6] := 0.000000e+000;
   STAT33[7, 10, 7] := 0.000000e+000;
   STAT33[7, 10, 8] := 0.000000e+000;
   STAT33[7, 10, 9] := 0.000000e+000;
   STAT33[7, 10, 10] := 0.000000e+000;
   STAT33[8, 1, 1] := 0.000000e+000;
   STAT33[8, 1, 2] := 0.000000e+000;
   STAT33[8, 1, 3] := 0.000000e+000;
   STAT33[8, 1, 4] := 0.000000e+000;
   STAT33[8, 1, 5] := 0.000000e+000;
   STAT33[8, 1, 6] := 0.000000e+000;
   STAT33[8, 1, 7] := 0.000000e+000;
   STAT33[8, 1, 8] := 0.000000e+000;
   STAT33[8, 1, 9] := 0.000000e+000;
   STAT33[8, 1, 10] := 0.000000e+000;
   STAT33[8, 2, 1] := 0.000000e+000;
   STAT33[8, 2, 2] := 0.000000e+000;
   STAT33[8, 2, 3] := 0.000000e+000;
   STAT33[8, 2, 4] := 0.000000e+000;
   STAT33[8, 2, 5] := 0.000000e+000;
   STAT33[8, 2, 6] := 0.000000e+000;
   STAT33[8, 2, 7] := 0.000000e+000;
   STAT33[8, 2, 8] := 0.000000e+000;
   STAT33[8, 2, 9] := 0.000000e+000;
   STAT33[8, 2, 10] := 0.000000e+000;
   STAT33[8, 3, 1] := 0.000000e+000;
   STAT33[8, 3, 2] := 0.000000e+000;
   STAT33[8, 3, 3] := 0.000000e+000;
   STAT33[8, 3, 4] := 0.000000e+000;
   STAT33[8, 3, 5] := 0.000000e+000;
   STAT33[8, 3, 6] := 0.000000e+000;
   STAT33[8, 3, 7] := 0.000000e+000;
   STAT33[8, 3, 8] := 0.000000e+000;
   STAT33[8, 3, 9] := 0.000000e+000;
   STAT33[8, 3, 10] := 0.000000e+000;
   STAT33[8, 4, 1] := 0.000000e+000;
   STAT33[8, 4, 2] := 0.000000e+000;
   STAT33[8, 4, 3] := 0.000000e+000;
   STAT33[8, 4, 4] := 0.000000e+000;
   STAT33[8, 4, 5] := 0.000000e+000;
   STAT33[8, 4, 6] := 0.000000e+000;
   STAT33[8, 4, 7] := 0.000000e+000;
   STAT33[8, 4, 8] := 0.000000e+000;
   STAT33[8, 4, 9] := 0.000000e+000;
   STAT33[8, 4, 10] := 0.000000e+000;
   STAT33[8, 5, 1] := 0.000000e+000;
   STAT33[8, 5, 2] := 0.000000e+000;
   STAT33[8, 5, 3] := 0.000000e+000;
   STAT33[8, 5, 4] := 0.000000e+000;
   STAT33[8, 5, 5] := 0.000000e+000;
   STAT33[8, 5, 6] := 0.000000e+000;
   STAT33[8, 5, 7] := 0.000000e+000;
   STAT33[8, 5, 8] := 0.000000e+000;
   STAT33[8, 5, 9] := 0.000000e+000;
   STAT33[8, 5, 10] := 0.000000e+000;
   STAT33[8, 6, 1] := 0.000000e+000;
   STAT33[8, 6, 2] := 0.000000e+000;
   STAT33[8, 6, 3] := 0.000000e+000;
   STAT33[8, 6, 4] := 0.000000e+000;
   STAT33[8, 6, 5] := 0.000000e+000;
   STAT33[8, 6, 6] := 0.000000e+000;
   STAT33[8, 6, 7] := 0.000000e+000;
   STAT33[8, 6, 8] := 0.000000e+000;
   STAT33[8, 6, 9] := 0.000000e+000;
   STAT33[8, 6, 10] := 0.000000e+000;
   STAT33[8, 7, 1] := 0.000000e+000;
   STAT33[8, 7, 2] := 0.000000e+000;
   STAT33[8, 7, 3] := 0.000000e+000;
   STAT33[8, 7, 4] := 0.000000e+000;
   STAT33[8, 7, 5] := 0.000000e+000;
   STAT33[8, 7, 6] := 0.000000e+000;
   STAT33[8, 7, 7] := 0.000000e+000;
   STAT33[8, 7, 8] := 0.000000e+000;
   STAT33[8, 7, 9] := 0.000000e+000;
   STAT33[8, 7, 10] := 0.000000e+000;
   STAT33[8, 8, 1] := 0.000000e+000;
   STAT33[8, 8, 2] := 0.000000e+000;
   STAT33[8, 8, 3] := 0.000000e+000;
   STAT33[8, 8, 4] := 0.000000e+000;
   STAT33[8, 8, 5] := 0.000000e+000;
   STAT33[8, 8, 6] := 0.000000e+000;
   STAT33[8, 8, 7] := 0.000000e+000;
   STAT33[8, 8, 8] := 0.000000e+000;
   STAT33[8, 8, 9] := 0.000000e+000;
   STAT33[8, 8, 10] := 0.000000e+000;
   STAT33[8, 9, 1] := 0.000000e+000;
   STAT33[8, 9, 2] := 0.000000e+000;
   STAT33[8, 9, 3] := 0.000000e+000;
   STAT33[8, 9, 4] := 0.000000e+000;
   STAT33[8, 9, 5] := 0.000000e+000;
   STAT33[8, 9, 6] := 0.000000e+000;
   STAT33[8, 9, 7] := 0.000000e+000;
   STAT33[8, 9, 8] := 0.000000e+000;
   STAT33[8, 9, 9] := 0.000000e+000;
   STAT33[8, 9, 10] := 0.000000e+000;
   STAT33[8, 10, 1] := 0.000000e+000;
   STAT33[8, 10, 2] := 0.000000e+000;
   STAT33[8, 10, 3] := 0.000000e+000;
   STAT33[8, 10, 4] := 0.000000e+000;
   STAT33[8, 10, 5] := 0.000000e+000;
   STAT33[8, 10, 6] := 0.000000e+000;
   STAT33[8, 10, 7] := 0.000000e+000;
   STAT33[8, 10, 8] := 0.000000e+000;
   STAT33[8, 10, 9] := 0.000000e+000;
   STAT33[8, 10, 10] := 0.000000e+000;
   STAT33[9, 1, 1] := 0.000000e+000;
   STAT33[9, 1, 2] := 0.000000e+000;
   STAT33[9, 1, 3] := 0.000000e+000;
   STAT33[9, 1, 4] := 0.000000e+000;
   STAT33[9, 1, 5] := 0.000000e+000;
   STAT33[9, 1, 6] := 0.000000e+000;
   STAT33[9, 1, 7] := 0.000000e+000;
   STAT33[9, 1, 8] := 0.000000e+000;
   STAT33[9, 1, 9] := 0.000000e+000;
   STAT33[9, 1, 10] := 0.000000e+000;
   STAT33[9, 2, 1] := 0.000000e+000;
   STAT33[9, 2, 2] := 0.000000e+000;
   STAT33[9, 2, 3] := 0.000000e+000;
   STAT33[9, 2, 4] := 0.000000e+000;
   STAT33[9, 2, 5] := 0.000000e+000;
   STAT33[9, 2, 6] := 0.000000e+000;
   STAT33[9, 2, 7] := 0.000000e+000;
   STAT33[9, 2, 8] := 0.000000e+000;
   STAT33[9, 2, 9] := 0.000000e+000;
   STAT33[9, 2, 10] := 0.000000e+000;
   STAT33[9, 3, 1] := 0.000000e+000;
   STAT33[9, 3, 2] := 0.000000e+000;
   STAT33[9, 3, 3] := 0.000000e+000;
   STAT33[9, 3, 4] := 0.000000e+000;
   STAT33[9, 3, 5] := 0.000000e+000;
   STAT33[9, 3, 6] := 0.000000e+000;
   STAT33[9, 3, 7] := 0.000000e+000;
   STAT33[9, 3, 8] := 0.000000e+000;
   STAT33[9, 3, 9] := 0.000000e+000;
   STAT33[9, 3, 10] := 0.000000e+000;
   STAT33[9, 4, 1] := 0.000000e+000;
   STAT33[9, 4, 2] := 0.000000e+000;
   STAT33[9, 4, 3] := 0.000000e+000;
   STAT33[9, 4, 4] := 0.000000e+000;
   STAT33[9, 4, 5] := 0.000000e+000;
   STAT33[9, 4, 6] := 0.000000e+000;
   STAT33[9, 4, 7] := 0.000000e+000;
   STAT33[9, 4, 8] := 0.000000e+000;
   STAT33[9, 4, 9] := 0.000000e+000;
   STAT33[9, 4, 10] := 0.000000e+000;
   STAT33[9, 5, 1] := 0.000000e+000;
   STAT33[9, 5, 2] := 0.000000e+000;
   STAT33[9, 5, 3] := 0.000000e+000;
   STAT33[9, 5, 4] := 0.000000e+000;
   STAT33[9, 5, 5] := 0.000000e+000;
   STAT33[9, 5, 6] := 0.000000e+000;
   STAT33[9, 5, 7] := 0.000000e+000;
   STAT33[9, 5, 8] := 0.000000e+000;
   STAT33[9, 5, 9] := 0.000000e+000;
   STAT33[9, 5, 10] := 0.000000e+000;
   STAT33[9, 6, 1] := 0.000000e+000;
   STAT33[9, 6, 2] := 0.000000e+000;
   STAT33[9, 6, 3] := 0.000000e+000;
   STAT33[9, 6, 4] := 0.000000e+000;
   STAT33[9, 6, 5] := 0.000000e+000;
   STAT33[9, 6, 6] := 0.000000e+000;
   STAT33[9, 6, 7] := 0.000000e+000;
   STAT33[9, 6, 8] := 0.000000e+000;
   STAT33[9, 6, 9] := 0.000000e+000;
   STAT33[9, 6, 10] := 0.000000e+000;
   STAT33[9, 7, 1] := 0.000000e+000;
   STAT33[9, 7, 2] := 0.000000e+000;
   STAT33[9, 7, 3] := 0.000000e+000;
   STAT33[9, 7, 4] := 0.000000e+000;
   STAT33[9, 7, 5] := 0.000000e+000;
   STAT33[9, 7, 6] := 0.000000e+000;
   STAT33[9, 7, 7] := 0.000000e+000;
   STAT33[9, 7, 8] := 0.000000e+000;
   STAT33[9, 7, 9] := 0.000000e+000;
   STAT33[9, 7, 10] := 0.000000e+000;
   STAT33[9, 8, 1] := 0.000000e+000;
   STAT33[9, 8, 2] := 0.000000e+000;
   STAT33[9, 8, 3] := 0.000000e+000;
   STAT33[9, 8, 4] := 0.000000e+000;
   STAT33[9, 8, 5] := 0.000000e+000;
   STAT33[9, 8, 6] := 0.000000e+000;
   STAT33[9, 8, 7] := 0.000000e+000;
   STAT33[9, 8, 8] := 0.000000e+000;
   STAT33[9, 8, 9] := 0.000000e+000;
   STAT33[9, 8, 10] := 0.000000e+000;
   STAT33[9, 9, 1] := 0.000000e+000;
   STAT33[9, 9, 2] := 0.000000e+000;
   STAT33[9, 9, 3] := 0.000000e+000;
   STAT33[9, 9, 4] := 0.000000e+000;
   STAT33[9, 9, 5] := 0.000000e+000;
   STAT33[9, 9, 6] := 0.000000e+000;
   STAT33[9, 9, 7] := 0.000000e+000;
   STAT33[9, 9, 8] := 0.000000e+000;
   STAT33[9, 9, 9] := 0.000000e+000;
   STAT33[9, 9, 10] := 0.000000e+000;
   STAT33[9, 10, 1] := 0.000000e+000;
   STAT33[9, 10, 2] := 0.000000e+000;
   STAT33[9, 10, 3] := 0.000000e+000;
   STAT33[9, 10, 4] := 0.000000e+000;
   STAT33[9, 10, 5] := 0.000000e+000;
   STAT33[9, 10, 6] := 0.000000e+000;
   STAT33[9, 10, 7] := 0.000000e+000;
   STAT33[9, 10, 8] := 0.000000e+000;
   STAT33[9, 10, 9] := 0.000000e+000;
   STAT33[9, 10, 10] := 0.000000e+000;
   STAT33[10, 1, 1] := 0.000000e+000;
   STAT33[10, 1, 2] := 0.000000e+000;
   STAT33[10, 1, 3] := 0.000000e+000;
   STAT33[10, 1, 4] := 0.000000e+000;
   STAT33[10, 1, 5] := 0.000000e+000;
   STAT33[10, 1, 6] := 0.000000e+000;
   STAT33[10, 1, 7] := 0.000000e+000;
   STAT33[10, 1, 8] := 0.000000e+000;
   STAT33[10, 1, 9] := 0.000000e+000;
   STAT33[10, 1, 10] := 0.000000e+000;
   STAT33[10, 2, 1] := 0.000000e+000;
   STAT33[10, 2, 2] := 0.000000e+000;
   STAT33[10, 2, 3] := 0.000000e+000;
   STAT33[10, 2, 4] := 0.000000e+000;
   STAT33[10, 2, 5] := 0.000000e+000;
   STAT33[10, 2, 6] := 0.000000e+000;
   STAT33[10, 2, 7] := 0.000000e+000;
   STAT33[10, 2, 8] := 0.000000e+000;
   STAT33[10, 2, 9] := 0.000000e+000;
   STAT33[10, 2, 10] := 0.000000e+000;
   STAT33[10, 3, 1] := 0.000000e+000;
   STAT33[10, 3, 2] := 0.000000e+000;
   STAT33[10, 3, 3] := 0.000000e+000;
   STAT33[10, 3, 4] := 0.000000e+000;
   STAT33[10, 3, 5] := 0.000000e+000;
   STAT33[10, 3, 6] := 0.000000e+000;
   STAT33[10, 3, 7] := 0.000000e+000;
   STAT33[10, 3, 8] := 0.000000e+000;
   STAT33[10, 3, 9] := 0.000000e+000;
   STAT33[10, 3, 10] := 0.000000e+000;
   STAT33[10, 4, 1] := 0.000000e+000;
   STAT33[10, 4, 2] := 0.000000e+000;
   STAT33[10, 4, 3] := 0.000000e+000;
   STAT33[10, 4, 4] := 0.000000e+000;
   STAT33[10, 4, 5] := 0.000000e+000;
   STAT33[10, 4, 6] := 0.000000e+000;
   STAT33[10, 4, 7] := 0.000000e+000;
   STAT33[10, 4, 8] := 0.000000e+000;
   STAT33[10, 4, 9] := 0.000000e+000;
   STAT33[10, 4, 10] := 0.000000e+000;
   STAT33[10, 5, 1] := 0.000000e+000;
   STAT33[10, 5, 2] := 0.000000e+000;
   STAT33[10, 5, 3] := 0.000000e+000;
   STAT33[10, 5, 4] := 0.000000e+000;
   STAT33[10, 5, 5] := 0.000000e+000;
   STAT33[10, 5, 6] := 0.000000e+000;
   STAT33[10, 5, 7] := 0.000000e+000;
   STAT33[10, 5, 8] := 0.000000e+000;
   STAT33[10, 5, 9] := 0.000000e+000;
   STAT33[10, 5, 10] := 0.000000e+000;
   STAT33[10, 6, 1] := 0.000000e+000;
   STAT33[10, 6, 2] := 0.000000e+000;
   STAT33[10, 6, 3] := 0.000000e+000;
   STAT33[10, 6, 4] := 0.000000e+000;
   STAT33[10, 6, 5] := 0.000000e+000;
   STAT33[10, 6, 6] := 0.000000e+000;
   STAT33[10, 6, 7] := 0.000000e+000;
   STAT33[10, 6, 8] := 0.000000e+000;
   STAT33[10, 6, 9] := 0.000000e+000;
   STAT33[10, 6, 10] := 0.000000e+000;
   STAT33[10, 7, 1] := 0.000000e+000;
   STAT33[10, 7, 2] := 0.000000e+000;
   STAT33[10, 7, 3] := 0.000000e+000;
   STAT33[10, 7, 4] := 0.000000e+000;
   STAT33[10, 7, 5] := 0.000000e+000;
   STAT33[10, 7, 6] := 0.000000e+000;
   STAT33[10, 7, 7] := 0.000000e+000;
   STAT33[10, 7, 8] := 0.000000e+000;
   STAT33[10, 7, 9] := 0.000000e+000;
   STAT33[10, 7, 10] := 0.000000e+000;
   STAT33[10, 8, 1] := 0.000000e+000;
   STAT33[10, 8, 2] := 0.000000e+000;
   STAT33[10, 8, 3] := 0.000000e+000;
   STAT33[10, 8, 4] := 0.000000e+000;
   STAT33[10, 8, 5] := 0.000000e+000;
   STAT33[10, 8, 6] := 0.000000e+000;
   STAT33[10, 8, 7] := 0.000000e+000;
   STAT33[10, 8, 8] := 0.000000e+000;
   STAT33[10, 8, 9] := 0.000000e+000;
   STAT33[10, 8, 10] := 0.000000e+000;
   STAT33[10, 9, 1] := 0.000000e+000;
   STAT33[10, 9, 2] := 0.000000e+000;
   STAT33[10, 9, 3] := 0.000000e+000;
   STAT33[10, 9, 4] := 0.000000e+000;
   STAT33[10, 9, 5] := 0.000000e+000;
   STAT33[10, 9, 6] := 0.000000e+000;
   STAT33[10, 9, 7] := 0.000000e+000;
   STAT33[10, 9, 8] := 0.000000e+000;
   STAT33[10, 9, 9] := 0.000000e+000;
   STAT33[10, 9, 10] := 0.000000e+000;
   STAT33[10, 10, 1] := 0.000000e+000;
   STAT33[10, 10, 2] := 0.000000e+000;
   STAT33[10, 10, 3] := 0.000000e+000;
   STAT33[10, 10, 4] := 0.000000e+000;
   STAT33[10, 10, 5] := 0.000000e+000;
   STAT33[10, 10, 6] := 0.000000e+000;
   STAT33[10, 10, 7] := 0.000000e+000;
   STAT33[10, 10, 8] := 0.000000e+000;
   STAT33[10, 10, 9] := 0.000000e+000;
   STAT33[10, 10, 10] := 0.000000e+000;
   STAT34[1] := 0;
   STAT34[2] := 0;
   STAT34[3] := 0;
   STAT34[4] := 0;
   STAT34[5] := 0;
   STAT34[6] := 0;
   STAT34[7] := 0;
   STAT34[8] := 0;
   STAT34[9] := 0;
   STAT34[10] := 0;
   STAT35[1] := FALSE;
   STAT35[2] := FALSE;
   STAT35[3] := FALSE;
   STAT35[4] := FALSE;
   STAT35[5] := FALSE;
   STAT35[6] := FALSE;
   STAT35[7] := FALSE;
   STAT35[8] := FALSE;
   STAT35[9] := FALSE;
   STAT35[10] := FALSE;
   STAT36[1] := FALSE;
   STAT36[2] := TRUE;
   STAT36[3] := TRUE;
   STAT36[4] := TRUE;
   STAT36[5] := TRUE;
   STAT36[6] := TRUE;
   STAT36[7] := TRUE;
   STAT36[8] := TRUE;
   STAT36[9] := TRUE;
   STAT36[10] := TRUE;
   STAT37[1] := FALSE;
   STAT37[2] := FALSE;
   STAT37[3] := FALSE;
   STAT37[4] := FALSE;
   STAT37[5] := FALSE;
   STAT37[6] := FALSE;
   STAT37[7] := FALSE;
   STAT37[8] := FALSE;
   STAT37[9] := FALSE;
   STAT37[10] := FALSE;
   STAT38[1].STAT39 := -5.394847e+003;
   STAT38[1].STAT40 := -1.542902e+003;
   STAT38[1].STAT41 := -2.054582e+003;
   STAT38[2].STAT39 := 8.890132e+002;
   STAT38[2].STAT40 := -1.497899e+003;
   STAT38[2].STAT41 := -2.149658e-001;
   STAT38[3].STAT39 := 8.919878e+002;
   STAT38[3].STAT40 := -1.090205e+003;
   STAT38[3].STAT41 := -9.505859e+000;
   STAT38[4].STAT39 := 8.918486e+002;
   STAT38[4].STAT40 := -2.388328e+003;
   STAT38[4].STAT41 := 1.638507e+003;
   STAT38[5].STAT39 := 0.000000e+000;
   STAT38[5].STAT40 := 0.000000e+000;
   STAT38[5].STAT41 := 0.000000e+000;
   STAT38[6].STAT39 := 0.000000e+000;
   STAT38[6].STAT40 := 0.000000e+000;
   STAT38[6].STAT41 := 0.000000e+000;
   STAT38[7].STAT39 := 0.000000e+000;
   STAT38[7].STAT40 := 0.000000e+000;
   STAT38[7].STAT41 := 0.000000e+000;
   STAT38[8].STAT39 := 0.000000e+000;
   STAT38[8].STAT40 := 0.000000e+000;
   STAT38[8].STAT41 := 0.000000e+000;
   STAT38[9].STAT39 := 0.000000e+000;
   STAT38[9].STAT40 := 0.000000e+000;
   STAT38[9].STAT41 := 0.000000e+000;
   STAT38[10].STAT39 := 0.000000e+000;
   STAT38[10].STAT40 := 0.000000e+000;
   STAT38[10].STAT41 := 0.000000e+000;
   STAT42[1].STAT43 := 1.692806e+004;
   STAT42[1].STAT44 := -7.794958e+003;
   STAT42[1].STAT45 := 1.076577e+004;
   STAT42[2].STAT43 := -7.713961e+003;
   STAT42[2].STAT44 := 4.273199e+003;
   STAT42[2].STAT45 := 1.898941e+004;
   STAT42[3].STAT43 := -2.348459e+003;
   STAT42[3].STAT44 := 7.782369e+003;
   STAT42[3].STAT45 := 1.453821e+004;
   STAT42[4].STAT43 := 5.917659e+003;
   STAT42[4].STAT44 := 1.137459e+004;
   STAT42[4].STAT45 := 3.265738e+004;
   STAT42[5].STAT43 := 0.000000e+000;
   STAT42[5].STAT44 := 0.000000e+000;
   STAT42[5].STAT45 := 0.000000e+000;
   STAT42[6].STAT43 := 0.000000e+000;
   STAT42[6].STAT44 := 0.000000e+000;
   STAT42[6].STAT45 := 0.000000e+000;
   STAT42[7].STAT43 := 0.000000e+000;
   STAT42[7].STAT44 := 0.000000e+000;
   STAT42[7].STAT45 := 0.000000e+000;
   STAT42[8].STAT43 := 0.000000e+000;
   STAT42[8].STAT44 := 0.000000e+000;
   STAT42[8].STAT45 := 0.000000e+000;
   STAT42[9].STAT43 := 0.000000e+000;
   STAT42[9].STAT44 := 0.000000e+000;
   STAT42[9].STAT45 := 0.000000e+000;
   STAT42[10].STAT43 := 0.000000e+000;
   STAT42[10].STAT44 := 0.000000e+000;
   STAT42[10].STAT45 := 0.000000e+000;
   STAT46 := 0;
   STAT47 := 0;
   STAT48[1].STAT49 := 0.000000e+000;
   STAT48[1].STAT50 := 0.000000e+000;
   STAT48[1].STAT51 := 0.000000e+000;
   STAT48[2].STAT49 := 0.000000e+000;
   STAT48[2].STAT50 := 0.000000e+000;
   STAT48[2].STAT51 := 0.000000e+000;
   STAT48[3].STAT49 := 0.000000e+000;
   STAT48[3].STAT50 := 0.000000e+000;
   STAT48[3].STAT51 := 0.000000e+000;
   STAT48[4].STAT49 := 0.000000e+000;
   STAT48[4].STAT50 := 0.000000e+000;
   STAT48[4].STAT51 := 0.000000e+000;
   STAT48[5].STAT49 := 0.000000e+000;
   STAT48[5].STAT50 := 0.000000e+000;
   STAT48[5].STAT51 := 0.000000e+000;
   STAT48[6].STAT49 := 0.000000e+000;
   STAT48[6].STAT50 := 0.000000e+000;
   STAT48[6].STAT51 := 0.000000e+000;
   STAT48[7].STAT49 := 0.000000e+000;
   STAT48[7].STAT50 := 0.000000e+000;
   STAT48[7].STAT51 := 0.000000e+000;
   STAT48[8].STAT49 := 0.000000e+000;
   STAT48[8].STAT50 := 0.000000e+000;
   STAT48[8].STAT51 := 0.000000e+000;
   STAT48[9].STAT49 := 0.000000e+000;
   STAT48[9].STAT50 := 0.000000e+000;
   STAT48[9].STAT51 := 0.000000e+000;
   STAT48[10].STAT49 := 0.000000e+000;
   STAT48[10].STAT50 := 0.000000e+000;
   STAT48[10].STAT51 := 0.000000e+000;
   STAT52[1].STAT53 := 0.000000e+000;
   STAT52[1].STAT54 := 0.000000e+000;
   STAT52[1].STAT55 := 0.000000e+000;
   STAT52[2].STAT53 := 0.000000e+000;
   STAT52[2].STAT54 := 0.000000e+000;
   STAT52[2].STAT55 := 0.000000e+000;
   STAT52[3].STAT53 := 0.000000e+000;
   STAT52[3].STAT54 := 0.000000e+000;
   STAT52[3].STAT55 := 0.000000e+000;
   STAT52[4].STAT53 := 0.000000e+000;
   STAT52[4].STAT54 := 0.000000e+000;
   STAT52[4].STAT55 := 0.000000e+000;
   STAT52[5].STAT53 := 0.000000e+000;
   STAT52[5].STAT54 := 0.000000e+000;
   STAT52[5].STAT55 := 0.000000e+000;
   STAT52[6].STAT53 := 0.000000e+000;
   STAT52[6].STAT54 := 0.000000e+000;
   STAT52[6].STAT55 := 0.000000e+000;
   STAT52[7].STAT53 := 0.000000e+000;
   STAT52[7].STAT54 := 0.000000e+000;
   STAT52[7].STAT55 := 0.000000e+000;
   STAT52[8].STAT53 := 0.000000e+000;
   STAT52[8].STAT54 := 0.000000e+000;
   STAT52[8].STAT55 := 0.000000e+000;
   STAT52[9].STAT53 := 0.000000e+000;
   STAT52[9].STAT54 := 0.000000e+000;
   STAT52[9].STAT55 := 0.000000e+000;
   STAT52[10].STAT53 := 0.000000e+000;
   STAT52[10].STAT54 := 0.000000e+000;
   STAT52[10].STAT55 := 0.000000e+000;
   STAT56 := 0;
   STAT57[1].STAT58 := -9.415735e+000;
   STAT57[1].STAT59 := -2.692465e+000;
   STAT57[1].STAT60 := -3.585904e+000;
   STAT57[2].STAT58 := 1.551612e+000;
   STAT57[2].STAT59 := -2.614949e+000;
   STAT57[2].STAT60 := -3.751841e-004;
   STAT57[3].STAT58 := 1.556804e+000;
   STAT57[3].STAT59 := -1.902676e+000;
   STAT57[3].STAT60 := -1.659077e-002;
   STAT57[4].STAT58 := 1.556561e+000;
   STAT57[4].STAT59 := -4.168549e+000;
   STAT57[4].STAT60 := 2.859719e+000;
   STAT57[5].STAT58 := 0.000000e+000;
   STAT57[5].STAT59 := 0.000000e+000;
   STAT57[5].STAT60 := 0.000000e+000;
   STAT57[6].STAT58 := 0.000000e+000;
   STAT57[6].STAT59 := 0.000000e+000;
   STAT57[6].STAT60 := 0.000000e+000;
   STAT57[7].STAT58 := 0.000000e+000;
   STAT57[7].STAT59 := 0.000000e+000;
   STAT57[7].STAT60 := 0.000000e+000;
   STAT57[8].STAT58 := 0.000000e+000;
   STAT57[8].STAT59 := 0.000000e+000;
   STAT57[8].STAT60 := 0.000000e+000;
   STAT57[9].STAT58 := 0.000000e+000;
   STAT57[9].STAT59 := 0.000000e+000;
   STAT57[9].STAT60 := 0.000000e+000;
   STAT57[10].STAT58 := 0.000000e+000;
   STAT57[10].STAT59 := 0.000000e+000;
   STAT57[10].STAT60 := 0.000000e+000;
   STAT61 := 0.000000e+000;
   STAT62 := 0.000000e+000;
   STAT63 := 0.000000e+000;
   STAT64[1].STAT65 := -4.147847e+003;
   STAT64[1].STAT66 := 7.063229e+002;
   STAT64[1].STAT67 := -2.065823e+002;
   STAT64[2].STAT65 := 2.161013e+003;
   STAT64[2].STAT66 := 2.477367e+002;
   STAT64[2].STAT67 := 1.742785e+003;
   STAT64[3].STAT65 := 2.158988e+003;
   STAT64[3].STAT66 := -1.661589e+002;
   STAT64[3].STAT67 := 3.479494e+003;
   STAT64[4].STAT65 := 2.147849e+003;
   STAT64[4].STAT66 := -2.054153e+002;
   STAT64[4].STAT67 := 3.480507e+003;
   STAT64[5].STAT65 := 0.000000e+000;
   STAT64[5].STAT66 := 0.000000e+000;
   STAT64[5].STAT67 := 0.000000e+000;
   STAT64[6].STAT65 := 0.000000e+000;
   STAT64[6].STAT66 := 0.000000e+000;
   STAT64[6].STAT67 := 0.000000e+000;
   STAT64[7].STAT65 := 0.000000e+000;
   STAT64[7].STAT66 := 0.000000e+000;
   STAT64[7].STAT67 := 0.000000e+000;
   STAT64[8].STAT65 := 0.000000e+000;
   STAT64[8].STAT66 := 0.000000e+000;
   STAT64[8].STAT67 := 0.000000e+000;
   STAT64[9].STAT65 := 0.000000e+000;
   STAT64[9].STAT66 := 0.000000e+000;
   STAT64[9].STAT67 := 0.000000e+000;
   STAT64[10].STAT65 := 0.000000e+000;
   STAT64[10].STAT66 := 0.000000e+000;
   STAT64[10].STAT67 := 0.000000e+000;
   STAT68 := FALSE;
   STAT69 := TRUE;
   STAT70 := FALSE;
   STAT71[1] := TRUE;
   STAT71[2] := FALSE;
   STAT71[3] := FALSE;
   STAT71[4] := FALSE;
   STAT71[5] := FALSE;
   STAT71[6] := FALSE;
   STAT71[7] := FALSE;
   STAT71[8] := FALSE;
   STAT71[9] := FALSE;
   STAT71[10] := FALSE;
END_DATA_BLOCK

DATA_BLOCK DB 23
VERSION : 0.0


  STRUCT
   STAT0 : INT ;
   STAT1 : REAL ;
   STAT2 : REAL ;
   STAT3 : REAL ;
   STAT4 : S5TIME ;
   STAT5 : ARRAY  [1 .. 10 ] OF STRUCT
    STAT6 : REAL ;
    STAT7 : REAL ;
   END_STRUCT ;
   STAT8 : REAL ;
   STAT9 : REAL ;
  END_STRUCT ;
BEGIN
   STAT0 := 50;
   STAT1 := 5.000000e+001;
   STAT2 := 5.000000e+001;
   STAT3 := 1.500000e+001;
   STAT4 := S5T#5S;
   STAT5[1].STAT6 := 0.000000e+000;
   STAT5[1].STAT7 := 0.000000e+000;
   STAT5[2].STAT6 := 4.000000e+003;
   STAT5[2].STAT7 := 0.000000e+000;
   STAT5[3].STAT6 := 8.000000e+003;
   STAT5[3].STAT7 := 0.000000e+000;
   STAT5[4].STAT6 := 1.200000e+004;
   STAT5[4].STAT7 := 0.000000e+000;
   STAT5[5].STAT6 := 0.000000e+000;
   STAT5[5].STAT7 := 0.000000e+000;
   STAT5[6].STAT6 := 0.000000e+000;
   STAT5[6].STAT7 := 0.000000e+000;
   STAT5[7].STAT6 := 0.000000e+000;
   STAT5[7].STAT7 := 0.000000e+000;
   STAT5[8].STAT6 := 0.000000e+000;
   STAT5[8].STAT7 := 0.000000e+000;
   STAT5[9].STAT6 := 0.000000e+000;
   STAT5[9].STAT7 := 0.000000e+000;
   STAT5[10].STAT6 := 0.000000e+000;
   STAT5[10].STAT7 := 0.000000e+000;
   STAT8 := 3.000000e+001;
   STAT9 := 1.000000e+002;
END_DATA_BLOCK

DATA_BLOCK DB 30
VERSION : 0.1


  STRUCT
   STAT0 : INT ;
   STAT1 : ARRAY  [1 .. 10 ] OF STRUCT
    STAT2 : DINT ;
    STAT3 : DINT ;
    STAT4 : DINT ;
   END_STRUCT ;
   STAT5 : INT ;
   STAT6 : INT ;
   STAT7 : INT ;
   STAT8 : INT ;
   STAT9 : ARRAY  [1 .. 10 ] OF STRUCT
    STAT10 : REAL ;
    STAT11 : REAL ;
    STAT12 : REAL ;
   END_STRUCT ;
   STAT13 : BOOL ;
   STAT14 : ARRAY  [1 .. 10 ] OF REAL ;
   STAT15 : ARRAY  [1 .. 10 ] OF REAL ;
   STAT16 : ARRAY  [1 .. 10 ] OF REAL ;
   STAT17 : ARRAY  [1 .. 10 ] OF REAL ;
   STAT18 : ARRAY  [1 .. 10 ] OF REAL ;
   STAT19 : ARRAY  [1 .. 10 ] OF REAL ;
   STAT20 : ARRAY  [1 .. 10 ] OF REAL ;
   STAT21 : BOOL  := TRUE;
   STAT22 : ARRAY  [1 .. 10 ] OF REAL ;
   STAT23 : ARRAY  [1 .. 10 ] OF REAL ;
   STAT24 : ARRAY  [1 .. 10 ] OF REAL ;
   STAT25 : ARRAY  [1 .. 10 ] OF REAL ;
   STAT26 : ARRAY  [1 .. 10 ] OF REAL ;
   STAT27 : ARRAY  [1 .. 10 ] OF REAL ;
   STAT28 : ARRAY  [1 .. 10 ] OF REAL ;
   STAT29 : BOOL ;
   STAT30 : ARRAY  [1 .. 10 ] OF STRUCT
    STAT31 : REAL ;
    STAT32 : REAL ;
    STAT33 : REAL ;
   END_STRUCT ;
   STAT34 : ARRAY  [1 .. 10 ] OF STRUCT
    STAT35 : REAL ;
    STAT36 : REAL ;
   END_STRUCT ;
  END_STRUCT ;
BEGIN
   STAT0 := 0;
   STAT1[1].STAT2 := L#884;
   STAT1[1].STAT3 := L#1006;
   STAT1[1].STAT4 := L#1770;
   STAT1[2].STAT2 := L#884;
   STAT1[2].STAT3 := L#1006;
   STAT1[2].STAT4 := L#1770;
   STAT1[3].STAT2 := L#884;
   STAT1[3].STAT3 := L#1006;
   STAT1[3].STAT4 := L#1770;
   STAT1[4].STAT2 := L#884;
   STAT1[4].STAT3 := L#1006;
   STAT1[4].STAT4 := L#1770;
   STAT1[5].STAT2 := L#0;
   STAT1[5].STAT3 := L#0;
   STAT1[5].STAT4 := L#0;
   STAT1[6].STAT2 := L#0;
   STAT1[6].STAT3 := L#0;
   STAT1[6].STAT4 := L#0;
   STAT1[7].STAT2 := L#0;
   STAT1[7].STAT3 := L#0;
   STAT1[7].STAT4 := L#0;
   STAT1[8].STAT2 := L#0;
   STAT1[8].STAT3 := L#0;
   STAT1[8].STAT4 := L#0;
   STAT1[9].STAT2 := L#0;
   STAT1[9].STAT3 := L#0;
   STAT1[9].STAT4 := L#0;
   STAT1[10].STAT2 := L#0;
   STAT1[10].STAT3 := L#0;
   STAT1[10].STAT4 := L#0;
   STAT5 := 50;
   STAT6 := 100;
   STAT7 := 600;
   STAT8 := 1000;
   STAT9[1].STAT10 := -1.247000e+003;
   STAT9[1].STAT11 := -2.249000e+003;
   STAT9[1].STAT12 := -1.848000e+003;
   STAT9[2].STAT10 := -1.272000e+003;
   STAT9[2].STAT11 := -1.746000e+003;
   STAT9[2].STAT12 := -1.743000e+003;
   STAT9[3].STAT10 := -1.267000e+003;
   STAT9[3].STAT11 := -9.240000e+002;
   STAT9[3].STAT12 := -3.489000e+003;
   STAT9[4].STAT10 := -1.256000e+003;
   STAT9[4].STAT11 := -2.183000e+003;
   STAT9[4].STAT12 := -1.842000e+003;
   STAT9[5].STAT10 := 0.000000e+000;
   STAT9[5].STAT11 := 0.000000e+000;
   STAT9[5].STAT12 := 0.000000e+000;
   STAT9[6].STAT10 := 0.000000e+000;
   STAT9[6].STAT11 := 0.000000e+000;
   STAT9[6].STAT12 := 0.000000e+000;
   STAT9[7].STAT10 := 0.000000e+000;
   STAT9[7].STAT11 := 0.000000e+000;
   STAT9[7].STAT12 := 0.000000e+000;
   STAT9[8].STAT10 := 0.000000e+000;
   STAT9[8].STAT11 := 0.000000e+000;
   STAT9[8].STAT12 := 0.000000e+000;
   STAT9[9].STAT10 := 0.000000e+000;
   STAT9[9].STAT11 := 0.000000e+000;
   STAT9[9].STAT12 := 0.000000e+000;
   STAT9[10].STAT10 := 0.000000e+000;
   STAT9[10].STAT11 := 0.000000e+000;
   STAT9[10].STAT12 := 0.000000e+000;
   STAT13 := TRUE;
   STAT14[1] := 2.064724e+000;
   STAT14[2] := 2.064724e+000;
   STAT14[3] := 2.064724e+000;
   STAT14[4] := 2.064724e+000;
   STAT14[5] := 0.000000e+000;
   STAT14[6] := 0.000000e+000;
   STAT14[7] := 0.000000e+000;
   STAT14[8] := 0.000000e+000;
   STAT14[9] := 0.000000e+000;
   STAT14[10] := 0.000000e+000;
   STAT15[1] := 5.585054e-001;
   STAT15[2] := 5.811946e-001;
   STAT15[3] := 1.919862e-001;
   STAT15[4] := 5.986480e-001;
   STAT15[5] := 0.000000e+000;
   STAT15[6] := 0.000000e+000;
   STAT15[7] := 0.000000e+000;
   STAT15[8] := 0.000000e+000;
   STAT15[9] := 0.000000e+000;
   STAT15[10] := 0.000000e+000;
   STAT16[1] := -3.839725e-001;
   STAT16[2] := -5.585054e-001;
   STAT16[3] := -5.811946e-001;
   STAT16[4] := -6.283185e-001;
   STAT16[5] := 0.000000e+000;
   STAT16[6] := 0.000000e+000;
   STAT16[7] := 0.000000e+000;
   STAT16[8] := 0.000000e+000;
   STAT16[9] := 0.000000e+000;
   STAT16[10] := 0.000000e+000;
   STAT17[1] := 0.000000e+000;
   STAT17[2] := 0.000000e+000;
   STAT17[3] := 0.000000e+000;
   STAT17[4] := 0.000000e+000;
   STAT17[5] := 0.000000e+000;
   STAT17[6] := 0.000000e+000;
   STAT17[7] := 0.000000e+000;
   STAT17[8] := 0.000000e+000;
   STAT17[9] := 0.000000e+000;
   STAT17[10] := 0.000000e+000;
   STAT18[1] := -3.490659e-001;
   STAT18[2] := -3.490659e-001;
   STAT18[3] := -3.490659e-001;
   STAT18[4] := -3.490659e-001;
   STAT18[5] := -2.268928e-001;
   STAT18[6] := -2.268928e-001;
   STAT18[7] := 0.000000e+000;
   STAT18[8] := 0.000000e+000;
   STAT18[9] := 0.000000e+000;
   STAT18[10] := 0.000000e+000;
   STAT19[1] := 8.726647e-002;
   STAT19[2] := 8.726647e-002;
   STAT19[3] := 8.726647e-002;
   STAT19[4] := 8.726647e-002;
   STAT19[5] := 0.000000e+000;
   STAT19[6] := 0.000000e+000;
   STAT19[7] := 0.000000e+000;
   STAT19[8] := 0.000000e+000;
   STAT19[9] := 0.000000e+000;
   STAT19[10] := 0.000000e+000;
   STAT20[1] := 0.000000e+000;
   STAT20[2] := 0.000000e+000;
   STAT20[3] := 0.000000e+000;
   STAT20[4] := 0.000000e+000;
   STAT20[5] := 0.000000e+000;
   STAT20[6] := 0.000000e+000;
   STAT20[7] := 0.000000e+000;
   STAT20[8] := 0.000000e+000;
   STAT20[9] := 0.000000e+000;
   STAT20[10] := 0.000000e+000;
   STAT21 := TRUE;
   STAT22[1] := 1.972222e+000;
   STAT22[2] := 1.972222e+000;
   STAT22[3] := 1.972222e+000;
   STAT22[4] := 1.972222e+000;
   STAT22[5] := 0.000000e+000;
   STAT22[6] := 0.000000e+000;
   STAT22[7] := 0.000000e+000;
   STAT22[8] := 0.000000e+000;
   STAT22[9] := 0.000000e+000;
   STAT22[10] := 0.000000e+000;
   STAT23[1] := 5.113815e-001;
   STAT23[2] := 5.410521e-001;
   STAT23[3] := 1.221731e-001;
   STAT23[4] := 5.462881e-001;
   STAT23[5] := 0.000000e+000;
   STAT23[6] := 0.000000e+000;
   STAT23[7] := 0.000000e+000;
   STAT23[8] := 0.000000e+000;
   STAT23[9] := 0.000000e+000;
   STAT23[10] := 0.000000e+000;
   STAT24[1] := -3.193952e-001;
   STAT24[2] := -5.061455e-001;
   STAT24[3] := -5.410521e-001;
   STAT24[4] := -5.811946e-001;
   STAT24[5] := 0.000000e+000;
   STAT24[6] := 0.000000e+000;
   STAT24[7] := 0.000000e+000;
   STAT24[8] := 0.000000e+000;
   STAT24[9] := 0.000000e+000;
   STAT24[10] := 0.000000e+000;
   STAT25[1] := 0.000000e+000;
   STAT25[2] := 0.000000e+000;
   STAT25[3] := 0.000000e+000;
   STAT25[4] := 0.000000e+000;
   STAT25[5] := 0.000000e+000;
   STAT25[6] := 0.000000e+000;
   STAT25[7] := 0.000000e+000;
   STAT25[8] := 0.000000e+000;
   STAT25[9] := 0.000000e+000;
   STAT25[10] := 0.000000e+000;
   STAT26[1] := -2.268928e-001;
   STAT26[2] := -2.268928e-001;
   STAT26[3] := -2.268928e-001;
   STAT26[4] := -2.268928e-001;
   STAT26[5] := 0.000000e+000;
   STAT26[6] := 0.000000e+000;
   STAT26[7] := 0.000000e+000;
   STAT26[8] := 0.000000e+000;
   STAT26[9] := 0.000000e+000;
   STAT26[10] := 0.000000e+000;
   STAT27[1] := -1.745329e-001;
   STAT27[2] := -1.745329e-001;
   STAT27[3] := -1.745329e-001;
   STAT27[4] := -1.745329e-001;
   STAT27[5] := -1.745329e-001;
   STAT27[6] := -1.745329e-001;
   STAT27[7] := 0.000000e+000;
   STAT27[8] := 0.000000e+000;
   STAT27[9] := 0.000000e+000;
   STAT27[10] := 0.000000e+000;
   STAT28[1] := 0.000000e+000;
   STAT28[2] := 0.000000e+000;
   STAT28[3] := 0.000000e+000;
   STAT28[4] := 0.000000e+000;
   STAT28[5] := 0.000000e+000;
   STAT28[6] := 0.000000e+000;
   STAT28[7] := 0.000000e+000;
   STAT28[8] := 0.000000e+000;
   STAT28[9] := 0.000000e+000;
   STAT28[10] := 0.000000e+000;
   STAT29 := FALSE;
   STAT30[1].STAT31 := 8.100000e+001;
   STAT30[1].STAT32 := -1.100000e+001;
   STAT30[1].STAT33 := -2.490000e+002;
   STAT30[2].STAT31 := 8.100000e+001;
   STAT30[2].STAT32 := -2.700000e+001;
   STAT30[2].STAT33 := -2.490000e+002;
   STAT30[3].STAT31 := 8.100000e+001;
   STAT30[3].STAT32 := 2.700000e+001;
   STAT30[3].STAT33 := -2.490000e+002;
   STAT30[4].STAT31 := 8.100000e+001;
   STAT30[4].STAT32 := 8.200000e+001;
   STAT30[4].STAT33 := -2.490000e+002;
   STAT30[5].STAT31 := 0.000000e+000;
   STAT30[5].STAT32 := 0.000000e+000;
   STAT30[5].STAT33 := 0.000000e+000;
   STAT30[6].STAT31 := 0.000000e+000;
   STAT30[6].STAT32 := 0.000000e+000;
   STAT30[6].STAT33 := 0.000000e+000;
   STAT30[7].STAT31 := 0.000000e+000;
   STAT30[7].STAT32 := 0.000000e+000;
   STAT30[7].STAT33 := 0.000000e+000;
   STAT30[8].STAT31 := 0.000000e+000;
   STAT30[8].STAT32 := 0.000000e+000;
   STAT30[8].STAT33 := 0.000000e+000;
   STAT30[9].STAT31 := 0.000000e+000;
   STAT30[9].STAT32 := 0.000000e+000;
   STAT30[9].STAT33 := 0.000000e+000;
   STAT30[10].STAT31 := 0.000000e+000;
   STAT30[10].STAT32 := 0.000000e+000;
   STAT30[10].STAT33 := 0.000000e+000;
   STAT34[1].STAT35 := 1.505000e+003;
   STAT34[1].STAT36 := 7.200000e+002;
   STAT34[2].STAT35 := 1.505000e+003;
   STAT34[2].STAT36 := 7.200000e+002;
   STAT34[3].STAT35 := 1.505000e+003;
   STAT34[3].STAT36 := 7.200000e+002;
   STAT34[4].STAT35 := 1.505000e+003;
   STAT34[4].STAT36 := 7.200000e+002;
   STAT34[5].STAT35 := 0.000000e+000;
   STAT34[5].STAT36 := 0.000000e+000;
   STAT34[6].STAT35 := 0.000000e+000;
   STAT34[6].STAT36 := 0.000000e+000;
   STAT34[7].STAT35 := 0.000000e+000;
   STAT34[7].STAT36 := 0.000000e+000;
   STAT34[8].STAT35 := 0.000000e+000;
   STAT34[8].STAT36 := 0.000000e+000;
   STAT34[9].STAT35 := 0.000000e+000;
   STAT34[9].STAT36 := 0.000000e+000;
   STAT34[10].STAT35 := 0.000000e+000;
   STAT34[10].STAT36 := 0.000000e+000;
END_DATA_BLOCK

DATA_BLOCK DB 50
VERSION : 0.1


  STRUCT
   STAT0 : ARRAY  [1 .. 64 ] OF BOOL ;
   STAT1 : ARRAY  [1 .. 6 ] OF WORD ;
   STAT2 : STRUCT
    STAT3 : BYTE ;
    STAT4 : BOOL ;
    STAT5 : BOOL ;
    STAT6 : BOOL ;
    STAT7 : BOOL ;
    STAT8 : BYTE ;
    STAT9 : BOOL ;
    STAT10 : BOOL ;
    STAT11 : BOOL ;
    STAT12 : BOOL ;
    STAT13 : BYTE ;
    STAT14 : BOOL ;
    STAT15 : BOOL ;
    STAT16 : BOOL ;
    STAT17 : BOOL ;
    STAT18 : ARRAY  [0 .. 3 ] OF BYTE ;
   END_STRUCT ;
   STAT19 : ARRAY  [1 .. 240 ] OF BOOL ;
   STAT20 : STRUCT
    STAT21 : INT ;
    STAT22 : WORD ;
    STAT23 : WORD ;
    STAT24 : INT ;
    STAT25 : WORD ;
    STAT26 : WORD ;
    STAT27 : WORD ;
    STAT28 : ARRAY  [1 .. 3 ] OF WORD ;
   END_STRUCT ;
   STAT29 : ARRAY  [1 .. 60 ] OF WORD ;
   STAT30 : ARRAY  [1 .. 240 ] OF BOOL ;
  END_STRUCT ;
BEGIN
   STAT0[1] := FALSE;
   STAT0[2] := FALSE;
   STAT0[3] := FALSE;
   STAT0[4] := FALSE;
   STAT0[5] := FALSE;
   STAT0[6] := FALSE;
   STAT0[7] := FALSE;
   STAT0[8] := TRUE;
   STAT0[9] := FALSE;
   STAT0[10] := FALSE;
   STAT0[11] := FALSE;
   STAT0[12] := FALSE;
   STAT0[13] := FALSE;
   STAT0[14] := FALSE;
   STAT0[15] := FALSE;
   STAT0[16] := FALSE;
   STAT0[17] := FALSE;
   STAT0[18] := FALSE;
   STAT0[19] := FALSE;
   STAT0[20] := FALSE;
   STAT0[21] := FALSE;
   STAT0[22] := FALSE;
   STAT0[23] := FALSE;
   STAT0[24] := FALSE;
   STAT0[25] := FALSE;
   STAT0[26] := FALSE;
   STAT0[27] := FALSE;
   STAT0[28] := FALSE;
   STAT0[29] := FALSE;
   STAT0[30] := FALSE;
   STAT0[31] := FALSE;
   STAT0[32] := FALSE;
   STAT0[33] := FALSE;
   STAT0[34] := FALSE;
   STAT0[35] := FALSE;
   STAT0[36] := FALSE;
   STAT0[37] := FALSE;
   STAT0[38] := FALSE;
   STAT0[39] := FALSE;
   STAT0[40] := FALSE;
   STAT0[41] := FALSE;
   STAT0[42] := FALSE;
   STAT0[43] := FALSE;
   STAT0[44] := FALSE;
   STAT0[45] := FALSE;
   STAT0[46] := FALSE;
   STAT0[47] := FALSE;
   STAT0[48] := FALSE;
   STAT0[49] := FALSE;
   STAT0[50] := FALSE;
   STAT0[51] := FALSE;
   STAT0[52] := FALSE;
   STAT0[53] := FALSE;
   STAT0[54] := FALSE;
   STAT0[55] := FALSE;
   STAT0[56] := FALSE;
   STAT0[57] := FALSE;
   STAT0[58] := FALSE;
   STAT0[59] := FALSE;
   STAT0[60] := FALSE;
   STAT0[61] := FALSE;
   STAT0[62] := FALSE;
   STAT0[63] := FALSE;
   STAT0[64] := FALSE;
   STAT1[1] := W#16#0;
   STAT1[2] := W#16#0;
   STAT1[3] := W#16#0;
   STAT1[4] := W#16#0;
   STAT1[5] := W#16#0;
   STAT1[6] := W#16#0;
   STAT2.STAT3 := B#16#0;
   STAT2.STAT4 := FALSE;
   STAT2.STAT5 := FALSE;
   STAT2.STAT6 := FALSE;
   STAT2.STAT7 := FALSE;
   STAT2.STAT8 := B#16#0;
   STAT2.STAT9 := FALSE;
   STAT2.STAT10 := TRUE;
   STAT2.STAT11 := FALSE;
   STAT2.STAT12 := FALSE;
   STAT2.STAT13 := B#16#0;
   STAT2.STAT14 := FALSE;
   STAT2.STAT15 := FALSE;
   STAT2.STAT16 := FALSE;
   STAT2.STAT17 := FALSE;
   STAT2.STAT18[0] := B#16#0;
   STAT2.STAT18[1] := B#16#0;
   STAT2.STAT18[2] := B#16#0;
   STAT2.STAT18[3] := B#16#0;
   STAT19[1] := FALSE;
   STAT19[2] := FALSE;
   STAT19[3] := FALSE;
   STAT19[4] := FALSE;
   STAT19[5] := FALSE;
   STAT19[6] := FALSE;
   STAT19[7] := FALSE;
   STAT19[8] := FALSE;
   STAT19[9] := FALSE;
   STAT19[10] := FALSE;
   STAT19[11] := FALSE;
   STAT19[12] := FALSE;
   STAT19[13] := FALSE;
   STAT19[14] := FALSE;
   STAT19[15] := FALSE;
   STAT19[16] := FALSE;
   STAT19[17] := FALSE;
   STAT19[18] := FALSE;
   STAT19[19] := FALSE;
   STAT19[20] := FALSE;
   STAT19[21] := FALSE;
   STAT19[22] := FALSE;
   STAT19[23] := FALSE;
   STAT19[24] := FALSE;
   STAT19[25] := FALSE;
   STAT19[26] := FALSE;
   STAT19[27] := FALSE;
   STAT19[28] := FALSE;
   STAT19[29] := FALSE;
   STAT19[30] := FALSE;
   STAT19[31] := FALSE;
   STAT19[32] := FALSE;
   STAT19[33] := FALSE;
   STAT19[34] := FALSE;
   STAT19[35] := FALSE;
   STAT19[36] := FALSE;
   STAT19[37] := FALSE;
   STAT19[38] := FALSE;
   STAT19[39] := FALSE;
   STAT19[40] := FALSE;
   STAT19[41] := FALSE;
   STAT19[42] := FALSE;
   STAT19[43] := FALSE;
   STAT19[44] := FALSE;
   STAT19[45] := FALSE;
   STAT19[46] := FALSE;
   STAT19[47] := FALSE;
   STAT19[48] := FALSE;
   STAT19[49] := FALSE;
   STAT19[50] := FALSE;
   STAT19[51] := FALSE;
   STAT19[52] := FALSE;
   STAT19[53] := FALSE;
   STAT19[54] := FALSE;
   STAT19[55] := FALSE;
   STAT19[56] := FALSE;
   STAT19[57] := FALSE;
   STAT19[58] := FALSE;
   STAT19[59] := FALSE;
   STAT19[60] := FALSE;
   STAT19[61] := FALSE;
   STAT19[62] := FALSE;
   STAT19[63] := FALSE;
   STAT19[64] := FALSE;
   STAT19[65] := FALSE;
   STAT19[66] := FALSE;
   STAT19[67] := FALSE;
   STAT19[68] := FALSE;
   STAT19[69] := FALSE;
   STAT19[70] := FALSE;
   STAT19[71] := FALSE;
   STAT19[72] := FALSE;
   STAT19[73] := FALSE;
   STAT19[74] := FALSE;
   STAT19[75] := FALSE;
   STAT19[76] := FALSE;
   STAT19[77] := FALSE;
   STAT19[78] := FALSE;
   STAT19[79] := FALSE;
   STAT19[80] := FALSE;
   STAT19[81] := FALSE;
   STAT19[82] := FALSE;
   STAT19[83] := FALSE;
   STAT19[84] := FALSE;
   STAT19[85] := FALSE;
   STAT19[86] := FALSE;
   STAT19[87] := FALSE;
   STAT19[88] := FALSE;
   STAT19[89] := FALSE;
   STAT19[90] := FALSE;
   STAT19[91] := FALSE;
   STAT19[92] := FALSE;
   STAT19[93] := FALSE;
   STAT19[94] := FALSE;
   STAT19[95] := FALSE;
   STAT19[96] := FALSE;
   STAT19[97] := FALSE;
   STAT19[98] := FALSE;
   STAT19[99] := FALSE;
   STAT19[100] := FALSE;
   STAT19[101] := FALSE;
   STAT19[102] := FALSE;
   STAT19[103] := FALSE;
   STAT19[104] := FALSE;
   STAT19[105] := FALSE;
   STAT19[106] := FALSE;
   STAT19[107] := FALSE;
   STAT19[108] := FALSE;
   STAT19[109] := FALSE;
   STAT19[110] := FALSE;
   STAT19[111] := FALSE;
   STAT19[112] := FALSE;
   STAT19[113] := FALSE;
   STAT19[114] := FALSE;
   STAT19[115] := FALSE;
   STAT19[116] := FALSE;
   STAT19[117] := FALSE;
   STAT19[118] := FALSE;
   STAT19[119] := FALSE;
   STAT19[120] := FALSE;
   STAT19[121] := FALSE;
   STAT19[122] := FALSE;
   STAT19[123] := FALSE;
   STAT19[124] := FALSE;
   STAT19[125] := FALSE;
   STAT19[126] := FALSE;
   STAT19[127] := FALSE;
   STAT19[128] := FALSE;
   STAT19[129] := FALSE;
   STAT19[130] := FALSE;
   STAT19[131] := FALSE;
   STAT19[132] := FALSE;
   STAT19[133] := FALSE;
   STAT19[134] := FALSE;
   STAT19[135] := FALSE;
   STAT19[136] := FALSE;
   STAT19[137] := FALSE;
   STAT19[138] := FALSE;
   STAT19[139] := FALSE;
   STAT19[140] := FALSE;
   STAT19[141] := FALSE;
   STAT19[142] := FALSE;
   STAT19[143] := FALSE;
   STAT19[144] := FALSE;
   STAT19[145] := FALSE;
   STAT19[146] := FALSE;
   STAT19[147] := FALSE;
   STAT19[148] := FALSE;
   STAT19[149] := FALSE;
   STAT19[150] := FALSE;
   STAT19[151] := FALSE;
   STAT19[152] := FALSE;
   STAT19[153] := FALSE;
   STAT19[154] := FALSE;
   STAT19[155] := FALSE;
   STAT19[156] := FALSE;
   STAT19[157] := FALSE;
   STAT19[158] := FALSE;
   STAT19[159] := FALSE;
   STAT19[160] := FALSE;
   STAT19[161] := FALSE;
   STAT19[162] := FALSE;
   STAT19[163] := FALSE;
   STAT19[164] := FALSE;
   STAT19[165] := FALSE;
   STAT19[166] := FALSE;
   STAT19[167] := FALSE;
   STAT19[168] := FALSE;
   STAT19[169] := FALSE;
   STAT19[170] := FALSE;
   STAT19[171] := FALSE;
   STAT19[172] := FALSE;
   STAT19[173] := FALSE;
   STAT19[174] := FALSE;
   STAT19[175] := FALSE;
   STAT19[176] := FALSE;
   STAT19[177] := FALSE;
   STAT19[178] := FALSE;
   STAT19[179] := FALSE;
   STAT19[180] := FALSE;
   STAT19[181] := FALSE;
   STAT19[182] := FALSE;
   STAT19[183] := FALSE;
   STAT19[184] := FALSE;
   STAT19[185] := FALSE;
   STAT19[186] := FALSE;
   STAT19[187] := FALSE;
   STAT19[188] := FALSE;
   STAT19[189] := FALSE;
   STAT19[190] := FALSE;
   STAT19[191] := FALSE;
   STAT19[192] := FALSE;
   STAT19[193] := FALSE;
   STAT19[194] := FALSE;
   STAT19[195] := FALSE;
   STAT19[196] := FALSE;
   STAT19[197] := FALSE;
   STAT19[198] := FALSE;
   STAT19[199] := FALSE;
   STAT19[200] := FALSE;
   STAT19[201] := FALSE;
   STAT19[202] := FALSE;
   STAT19[203] := FALSE;
   STAT19[204] := FALSE;
   STAT19[205] := FALSE;
   STAT19[206] := FALSE;
   STAT19[207] := FALSE;
   STAT19[208] := FALSE;
   STAT19[209] := FALSE;
   STAT19[210] := FALSE;
   STAT19[211] := FALSE;
   STAT19[212] := FALSE;
   STAT19[213] := FALSE;
   STAT19[214] := FALSE;
   STAT19[215] := FALSE;
   STAT19[216] := FALSE;
   STAT19[217] := FALSE;
   STAT19[218] := FALSE;
   STAT19[219] := FALSE;
   STAT19[220] := FALSE;
   STAT19[221] := FALSE;
   STAT19[222] := FALSE;
   STAT19[223] := FALSE;
   STAT19[224] := FALSE;
   STAT19[225] := FALSE;
   STAT19[226] := FALSE;
   STAT19[227] := FALSE;
   STAT19[228] := FALSE;
   STAT19[229] := FALSE;
   STAT19[230] := FALSE;
   STAT19[231] := FALSE;
   STAT19[232] := FALSE;
   STAT19[233] := FALSE;
   STAT19[234] := FALSE;
   STAT19[235] := FALSE;
   STAT19[236] := FALSE;
   STAT19[237] := FALSE;
   STAT19[238] := FALSE;
   STAT19[239] := FALSE;
   STAT19[240] := FALSE;
   STAT20.STAT21 := 0;
   STAT20.STAT22 := W#16#0;
   STAT20.STAT23 := W#16#0;
   STAT20.STAT24 := 0;
   STAT20.STAT25 := W#16#0;
   STAT20.STAT26 := W#16#0;
   STAT20.STAT27 := W#16#0;
   STAT20.STAT28[1] := W#16#0;
   STAT20.STAT28[2] := W#16#0;
   STAT20.STAT28[3] := W#16#0;
   STAT29[1] := W#16#0;
   STAT29[2] := W#16#0;
   STAT29[3] := W#16#0;
   STAT29[4] := W#16#0;
   STAT29[5] := W#16#0;
   STAT29[6] := W#16#0;
   STAT29[7] := W#16#0;
   STAT29[8] := W#16#0;
   STAT29[9] := W#16#0;
   STAT29[10] := W#16#0;
   STAT29[11] := W#16#0;
   STAT29[12] := W#16#0;
   STAT29[13] := W#16#0;
   STAT29[14] := W#16#0;
   STAT29[15] := W#16#0;
   STAT29[16] := W#16#0;
   STAT29[17] := W#16#0;
   STAT29[18] := W#16#0;
   STAT29[19] := W#16#0;
   STAT29[20] := W#16#0;
   STAT29[21] := W#16#0;
   STAT29[22] := W#16#0;
   STAT29[23] := W#16#0;
   STAT29[24] := W#16#0;
   STAT29[25] := W#16#0;
   STAT29[26] := W#16#0;
   STAT29[27] := W#16#0;
   STAT29[28] := W#16#0;
   STAT29[29] := W#16#0;
   STAT29[30] := W#16#0;
   STAT29[31] := W#16#0;
   STAT29[32] := W#16#0;
   STAT29[33] := W#16#0;
   STAT29[34] := W#16#0;
   STAT29[35] := W#16#0;
   STAT29[36] := W#16#0;
   STAT29[37] := W#16#0;
   STAT29[38] := W#16#0;
   STAT29[39] := W#16#0;
   STAT29[40] := W#16#0;
   STAT29[41] := W#16#0;
   STAT29[42] := W#16#0;
   STAT29[43] := W#16#0;
   STAT29[44] := W#16#0;
   STAT29[45] := W#16#0;
   STAT29[46] := W#16#0;
   STAT29[47] := W#16#0;
   STAT29[48] := W#16#0;
   STAT29[49] := W#16#0;
   STAT29[50] := W#16#0;
   STAT29[51] := W#16#0;
   STAT29[52] := W#16#0;
   STAT29[53] := W#16#0;
   STAT29[54] := W#16#0;
   STAT29[55] := W#16#0;
   STAT29[56] := W#16#0;
   STAT29[57] := W#16#0;
   STAT29[58] := W#16#0;
   STAT29[59] := W#16#0;
   STAT29[60] := W#16#0;
   STAT30[1] := FALSE;
   STAT30[2] := FALSE;
   STAT30[3] := FALSE;
   STAT30[4] := FALSE;
   STAT30[5] := FALSE;
   STAT30[6] := FALSE;
   STAT30[7] := FALSE;
   STAT30[8] := FALSE;
   STAT30[9] := FALSE;
   STAT30[10] := FALSE;
   STAT30[11] := FALSE;
   STAT30[12] := FALSE;
   STAT30[13] := FALSE;
   STAT30[14] := FALSE;
   STAT30[15] := FALSE;
   STAT30[16] := FALSE;
   STAT30[17] := FALSE;
   STAT30[18] := FALSE;
   STAT30[19] := FALSE;
   STAT30[20] := FALSE;
   STAT30[21] := FALSE;
   STAT30[22] := FALSE;
   STAT30[23] := FALSE;
   STAT30[24] := FALSE;
   STAT30[25] := FALSE;
   STAT30[26] := FALSE;
   STAT30[27] := FALSE;
   STAT30[28] := FALSE;
   STAT30[29] := FALSE;
   STAT30[30] := FALSE;
   STAT30[31] := FALSE;
   STAT30[32] := FALSE;
   STAT30[33] := FALSE;
   STAT30[34] := FALSE;
   STAT30[35] := FALSE;
   STAT30[36] := FALSE;
   STAT30[37] := FALSE;
   STAT30[38] := FALSE;
   STAT30[39] := FALSE;
   STAT30[40] := FALSE;
   STAT30[41] := FALSE;
   STAT30[42] := FALSE;
   STAT30[43] := FALSE;
   STAT30[44] := FALSE;
   STAT30[45] := FALSE;
   STAT30[46] := FALSE;
   STAT30[47] := FALSE;
   STAT30[48] := FALSE;
   STAT30[49] := FALSE;
   STAT30[50] := FALSE;
   STAT30[51] := FALSE;
   STAT30[52] := FALSE;
   STAT30[53] := FALSE;
   STAT30[54] := FALSE;
   STAT30[55] := FALSE;
   STAT30[56] := FALSE;
   STAT30[57] := FALSE;
   STAT30[58] := FALSE;
   STAT30[59] := FALSE;
   STAT30[60] := FALSE;
   STAT30[61] := FALSE;
   STAT30[62] := FALSE;
   STAT30[63] := FALSE;
   STAT30[64] := FALSE;
   STAT30[65] := FALSE;
   STAT30[66] := FALSE;
   STAT30[67] := FALSE;
   STAT30[68] := FALSE;
   STAT30[69] := FALSE;
   STAT30[70] := FALSE;
   STAT30[71] := FALSE;
   STAT30[72] := FALSE;
   STAT30[73] := FALSE;
   STAT30[74] := FALSE;
   STAT30[75] := FALSE;
   STAT30[76] := FALSE;
   STAT30[77] := FALSE;
   STAT30[78] := FALSE;
   STAT30[79] := FALSE;
   STAT30[80] := FALSE;
   STAT30[81] := FALSE;
   STAT30[82] := FALSE;
   STAT30[83] := FALSE;
   STAT30[84] := FALSE;
   STAT30[85] := FALSE;
   STAT30[86] := FALSE;
   STAT30[87] := FALSE;
   STAT30[88] := FALSE;
   STAT30[89] := FALSE;
   STAT30[90] := FALSE;
   STAT30[91] := FALSE;
   STAT30[92] := FALSE;
   STAT30[93] := FALSE;
   STAT30[94] := FALSE;
   STAT30[95] := FALSE;
   STAT30[96] := FALSE;
   STAT30[97] := FALSE;
   STAT30[98] := FALSE;
   STAT30[99] := FALSE;
   STAT30[100] := FALSE;
   STAT30[101] := FALSE;
   STAT30[102] := FALSE;
   STAT30[103] := FALSE;
   STAT30[104] := FALSE;
   STAT30[105] := FALSE;
   STAT30[106] := FALSE;
   STAT30[107] := FALSE;
   STAT30[108] := FALSE;
   STAT30[109] := FALSE;
   STAT30[110] := FALSE;
   STAT30[111] := FALSE;
   STAT30[112] := FALSE;
   STAT30[113] := FALSE;
   STAT30[114] := FALSE;
   STAT30[115] := FALSE;
   STAT30[116] := FALSE;
   STAT30[117] := FALSE;
   STAT30[118] := FALSE;
   STAT30[119] := FALSE;
   STAT30[120] := FALSE;
   STAT30[121] := FALSE;
   STAT30[122] := FALSE;
   STAT30[123] := FALSE;
   STAT30[124] := FALSE;
   STAT30[125] := FALSE;
   STAT30[126] := FALSE;
   STAT30[127] := FALSE;
   STAT30[128] := FALSE;
   STAT30[129] := FALSE;
   STAT30[130] := FALSE;
   STAT30[131] := FALSE;
   STAT30[132] := FALSE;
   STAT30[133] := FALSE;
   STAT30[134] := FALSE;
   STAT30[135] := FALSE;
   STAT30[136] := FALSE;
   STAT30[137] := FALSE;
   STAT30[138] := FALSE;
   STAT30[139] := FALSE;
   STAT30[140] := FALSE;
   STAT30[141] := FALSE;
   STAT30[142] := FALSE;
   STAT30[143] := FALSE;
   STAT30[144] := FALSE;
   STAT30[145] := FALSE;
   STAT30[146] := FALSE;
   STAT30[147] := FALSE;
   STAT30[148] := FALSE;
   STAT30[149] := FALSE;
   STAT30[150] := FALSE;
   STAT30[151] := FALSE;
   STAT30[152] := FALSE;
   STAT30[153] := FALSE;
   STAT30[154] := FALSE;
   STAT30[155] := FALSE;
   STAT30[156] := FALSE;
   STAT30[157] := FALSE;
   STAT30[158] := FALSE;
   STAT30[159] := FALSE;
   STAT30[160] := FALSE;
   STAT30[161] := FALSE;
   STAT30[162] := FALSE;
   STAT30[163] := FALSE;
   STAT30[164] := FALSE;
   STAT30[165] := FALSE;
   STAT30[166] := FALSE;
   STAT30[167] := FALSE;
   STAT30[168] := FALSE;
   STAT30[169] := FALSE;
   STAT30[170] := FALSE;
   STAT30[171] := FALSE;
   STAT30[172] := FALSE;
   STAT30[173] := FALSE;
   STAT30[174] := FALSE;
   STAT30[175] := FALSE;
   STAT30[176] := FALSE;
   STAT30[177] := FALSE;
   STAT30[178] := FALSE;
   STAT30[179] := FALSE;
   STAT30[180] := FALSE;
   STAT30[181] := FALSE;
   STAT30[182] := FALSE;
   STAT30[183] := FALSE;
   STAT30[184] := FALSE;
   STAT30[185] := FALSE;
   STAT30[186] := FALSE;
   STAT30[187] := FALSE;
   STAT30[188] := FALSE;
   STAT30[189] := FALSE;
   STAT30[190] := FALSE;
   STAT30[191] := FALSE;
   STAT30[192] := FALSE;
   STAT30[193] := FALSE;
   STAT30[194] := FALSE;
   STAT30[195] := FALSE;
   STAT30[196] := FALSE;
   STAT30[197] := FALSE;
   STAT30[198] := FALSE;
   STAT30[199] := FALSE;
   STAT30[200] := FALSE;
   STAT30[201] := FALSE;
   STAT30[202] := FALSE;
   STAT30[203] := FALSE;
   STAT30[204] := FALSE;
   STAT30[205] := FALSE;
   STAT30[206] := FALSE;
   STAT30[207] := FALSE;
   STAT30[208] := FALSE;
   STAT30[209] := FALSE;
   STAT30[210] := FALSE;
   STAT30[211] := FALSE;
   STAT30[212] := FALSE;
   STAT30[213] := FALSE;
   STAT30[214] := FALSE;
   STAT30[215] := FALSE;
   STAT30[216] := FALSE;
   STAT30[217] := FALSE;
   STAT30[218] := FALSE;
   STAT30[219] := FALSE;
   STAT30[220] := FALSE;
   STAT30[221] := FALSE;
   STAT30[222] := FALSE;
   STAT30[223] := FALSE;
   STAT30[224] := FALSE;
   STAT30[225] := FALSE;
   STAT30[226] := FALSE;
   STAT30[227] := FALSE;
   STAT30[228] := FALSE;
   STAT30[229] := FALSE;
   STAT30[230] := FALSE;
   STAT30[231] := FALSE;
   STAT30[232] := FALSE;
   STAT30[233] := FALSE;
   STAT30[234] := FALSE;
   STAT30[235] := FALSE;
   STAT30[236] := FALSE;
   STAT30[237] := FALSE;
   STAT30[238] := FALSE;
   STAT30[239] := FALSE;
   STAT30[240] := FALSE;
END_DATA_BLOCK

DATA_BLOCK DB 51
VERSION : 0.1


  STRUCT
   STAT0 : BOOL ;
   STAT1 : BOOL ;
   STAT2 : BOOL ;
   STAT3 : BOOL ;
   STAT4 : BOOL ;
   STAT5 : BOOL ;
   STAT6 : BOOL ;
   STAT7 : ARRAY  [1 .. 10 ] OF BOOL ;
   STAT8 : ARRAY  [1 .. 10 ] OF BOOL ;
   STAT9 : ARRAY  [1 .. 10 ] OF BOOL ;
   STAT10 : ARRAY  [1 .. 10 ] OF BOOL ;
   STAT11 : ARRAY  [1 .. 10 ] OF BOOL ;
   STAT12 : ARRAY  [1 .. 10 ] OF REAL ;
   STAT13 : ARRAY  [1 .. 10 ] OF REAL ;
   STAT14 : ARRAY  [1 .. 10 ] OF REAL ;
   STAT15 : ARRAY  [1 .. 10 ] OF REAL ;
   STAT16 : ARRAY  [1 .. 10 ] OF REAL ;
   STAT17 : ARRAY  [1 .. 10 ] OF REAL ;
   STAT18 : ARRAY  [1 .. 10 ] OF REAL ;
   STAT19 : ARRAY  [1 .. 10 ] OF REAL ;
   STAT20 : INT ;
   STAT21 : INT ;
   STAT22 : INT ;
   STAT23 : INT ;
   STAT24 : INT ;
   STAT25 : REAL ;
   STAT26 : REAL ;
   STAT27 : REAL ;
   STAT28 : REAL ;
   STAT29 : REAL ;
   STAT30 : REAL ;
   STAT31 : REAL ;
   STAT32 : REAL ;
   STAT33 : INT ;
   STAT34 : INT ;
   STAT35 : INT ;
   STAT36 : INT ;
   STAT37 : INT ;
   STAT38 : INT ;
  END_STRUCT ;
BEGIN
   STAT0 := FALSE;
   STAT1 := TRUE;
   STAT2 := FALSE;
   STAT3 := FALSE;
   STAT4 := FALSE;
   STAT5 := FALSE;
   STAT6 := FALSE;
   STAT7[1] := FALSE;
   STAT7[2] := FALSE;
   STAT7[3] := FALSE;
   STAT7[4] := FALSE;
   STAT7[5] := FALSE;
   STAT7[6] := FALSE;
   STAT7[7] := FALSE;
   STAT7[8] := FALSE;
   STAT7[9] := FALSE;
   STAT7[10] := FALSE;
   STAT8[1] := FALSE;
   STAT8[2] := FALSE;
   STAT8[3] := FALSE;
   STAT8[4] := FALSE;
   STAT8[5] := FALSE;
   STAT8[6] := FALSE;
   STAT8[7] := FALSE;
   STAT8[8] := FALSE;
   STAT8[9] := FALSE;
   STAT8[10] := FALSE;
   STAT9[1] := FALSE;
   STAT9[2] := FALSE;
   STAT9[3] := FALSE;
   STAT9[4] := FALSE;
   STAT9[5] := FALSE;
   STAT9[6] := FALSE;
   STAT9[7] := FALSE;
   STAT9[8] := FALSE;
   STAT9[9] := FALSE;
   STAT9[10] := FALSE;
   STAT10[1] := FALSE;
   STAT10[2] := FALSE;
   STAT10[3] := FALSE;
   STAT10[4] := FALSE;
   STAT10[5] := FALSE;
   STAT10[6] := FALSE;
   STAT10[7] := FALSE;
   STAT10[8] := FALSE;
   STAT10[9] := FALSE;
   STAT10[10] := FALSE;
   STAT11[1] := TRUE;
   STAT11[2] := FALSE;
   STAT11[3] := FALSE;
   STAT11[4] := FALSE;
   STAT11[5] := FALSE;
   STAT11[6] := FALSE;
   STAT11[7] := FALSE;
   STAT11[8] := FALSE;
   STAT11[9] := FALSE;
   STAT11[10] := FALSE;
   STAT12[1] := -3.132479e+000;
   STAT12[2] := 2.384183e+001;
   STAT12[3] := 1.891271e+001;
   STAT12[4] := 1.#QNAN0e+000;
   STAT12[5] := 0.000000e+000;
   STAT12[6] := 0.000000e+000;
   STAT12[7] := 0.000000e+000;
   STAT12[8] := 0.000000e+000;
   STAT12[9] := 0.000000e+000;
   STAT12[10] := 0.000000e+000;
   STAT13[1] := -2.580451e+000;
   STAT13[2] := -4.761978e+000;
   STAT13[3] := -1.799458e+000;
   STAT13[4] := 3.709789e+000;
   STAT13[5] := 0.000000e+000;
   STAT13[6] := 0.000000e+000;
   STAT13[7] := 0.000000e+000;
   STAT13[8] := 0.000000e+000;
   STAT13[9] := 0.000000e+000;
   STAT13[10] := 0.000000e+000;
   STAT14[1] := 1.696736e+001;
   STAT14[2] := -5.081615e+000;
   STAT14[3] := -4.419737e-001;
   STAT14[4] := 2.768813e+000;
   STAT14[5] := 0.000000e+000;
   STAT14[6] := 0.000000e+000;
   STAT14[7] := 0.000000e+000;
   STAT14[8] := 0.000000e+000;
   STAT14[9] := 0.000000e+000;
   STAT14[10] := 0.000000e+000;
   STAT15[1] := -2.575637e+000;
   STAT15[2] := 2.431845e+001;
   STAT15[3] := 1.937624e+001;
   STAT15[4] := 1.#QNAN0e+000;
   STAT15[5] := 0.000000e+000;
   STAT15[6] := 0.000000e+000;
   STAT15[7] := 0.000000e+000;
   STAT15[8] := 0.000000e+000;
   STAT15[9] := 0.000000e+000;
   STAT15[10] := 0.000000e+000;
   STAT16[1] := -1.401561e+000;
   STAT16[2] := -5.373302e+000;
   STAT16[3] := -1.968241e+000;
   STAT16[4] := 4.097909e+000;
   STAT16[5] := 0.000000e+000;
   STAT16[6] := 0.000000e+000;
   STAT16[7] := 0.000000e+000;
   STAT16[8] := 0.000000e+000;
   STAT16[9] := 0.000000e+000;
   STAT16[10] := 0.000000e+000;
   STAT17[1] := 1.799781e+001;
   STAT17[2] := -5.550834e+000;
   STAT17[3] := -6.710100e-001;
   STAT17[4] := 3.114355e+000;
   STAT17[5] := 0.000000e+000;
   STAT17[6] := 0.000000e+000;
   STAT17[7] := 0.000000e+000;
   STAT17[8] := 0.000000e+000;
   STAT17[9] := 0.000000e+000;
   STAT17[10] := 0.000000e+000;
   STAT18[1] := 4.281171e+000;
   STAT18[2] := -3.940207e+000;
   STAT18[3] := 5.123652e-001;
   STAT18[4] := -1.760909e+001;
   STAT18[5] := 0.000000e+000;
   STAT18[6] := 0.000000e+000;
   STAT18[7] := 0.000000e+000;
   STAT18[8] := 0.000000e+000;
   STAT18[9] := 0.000000e+000;
   STAT18[10] := 0.000000e+000;
   STAT19[1] := 3.568829e+000;
   STAT19[2] := 1.179021e+001;
   STAT19[3] := 7.337635e+000;
   STAT19[4] := 2.545909e+001;
   STAT19[5] := 0.000000e+000;
   STAT19[6] := 0.000000e+000;
   STAT19[7] := 0.000000e+000;
   STAT19[8] := 0.000000e+000;
   STAT19[9] := 0.000000e+000;
   STAT19[10] := 0.000000e+000;
   STAT20 := -10;
   STAT21 := -10;
   STAT22 := -10;
   STAT23 := -10;
   STAT24 := -10;
   STAT25 := 0.000000e+000;
   STAT26 := 0.000000e+000;
   STAT27 := 0.000000e+000;
   STAT28 := 0.000000e+000;
   STAT29 := 0.000000e+000;
   STAT30 := 0.000000e+000;
   STAT31 := 0.000000e+000;
   STAT32 := 0.000000e+000;
   STAT33 := 0;
   STAT34 := 0;
   STAT35 := 0;
   STAT36 := 0;
   STAT37 := 0;
   STAT38 := 0;
END_DATA_BLOCK

DATA_BLOCK DB 95
VERSION : 0.1


  STRUCT
   STAT0 : STRUCT
    STAT1 : BOOL ;
    STAT2 : BOOL ;
    STAT3 : BOOL ;
    STAT4 : BOOL ;
    STAT5 : BOOL ;
    STAT6 : BOOL ;
    STAT7 : BOOL ;
    STAT8 : BOOL ;
    STAT9 : BOOL ;
    STAT10 : BOOL ;
    STAT11 : BOOL ;
    STAT12 : BOOL ;
    STAT13 : BOOL ;
    STAT14 : BOOL ;
    STAT15 : BOOL ;
    STAT16 : BOOL ;
    STAT17 : ARRAY  [0 .. 7 ] OF WORD ;
   END_STRUCT ;
   STAT18 : STRUCT
    STAT19 : INT ;
    STAT20 : INT ;
    STAT21 : INT ;
    STAT22 : INT ;
    STAT23 : INT ;
    STAT24 : INT ;
    STAT25 : INT ;
    STAT26 : INT ;
    STAT27 : INT ;
    STAT28 : INT ;
   END_STRUCT ;
   STAT29 : STRUCT
    STAT30 : INT ;
    STAT31 : INT ;
    STAT32 : INT ;
    STAT33 : INT ;
    STAT34 : INT ;
    STAT35 : INT ;
    STAT36 : INT ;
    STAT37 : INT ;
    STAT38 : INT ;
    STAT39 : INT ;
   END_STRUCT ;
   STAT40 : STRUCT
    STAT41 : INT ;
    STAT42 : INT ;
    STAT43 : INT ;
    STAT44 : INT ;
    STAT45 : INT ;
    STAT46 : INT ;
    STAT47 : INT ;
    STAT48 : INT ;
    STAT49 : INT ;
    STAT50 : INT ;
   END_STRUCT ;
   STAT51 : STRUCT
    STAT52 : INT ;
    STAT53 : INT ;
    STAT54 : INT ;
    STAT55 : INT ;
    STAT56 : INT ;
    STAT57 : INT ;
    STAT58 : INT ;
    STAT59 : INT ;
    STAT60 : INT ;
    STAT61 : INT ;
   END_STRUCT ;
   STAT62 : STRUCT
    STAT63 : INT ;
    STAT64 : INT ;
    STAT65 : INT ;
    STAT66 : INT ;
    STAT67 : INT ;
    STAT68 : INT ;
    STAT69 : INT ;
    STAT70 : INT ;
    STAT71 : INT ;
    STAT72 : INT ;
   END_STRUCT ;
   STAT73 : STRUCT
    STAT74 : INT ;
    STAT75 : INT ;
    STAT76 : INT ;
    STAT77 : INT ;
    STAT78 : INT ;
    STAT79 : INT ;
    STAT80 : INT ;
    STAT81 : INT ;
    STAT82 : INT ;
    STAT83 : INT ;
   END_STRUCT ;
   STAT84 : STRUCT
    STAT85 : INT ;
    STAT86 : INT ;
    STAT87 : INT ;
    STAT88 : INT ;
    STAT89 : INT ;
    STAT90 : INT ;
    STAT91 : INT ;
    STAT92 : INT ;
    STAT93 : INT ;
    STAT94 : INT ;
   END_STRUCT ;
  END_STRUCT ;
BEGIN
   STAT0.STAT1 := FALSE;
   STAT0.STAT2 := FALSE;
   STAT0.STAT3 := FALSE;
   STAT0.STAT4 := FALSE;
   STAT0.STAT5 := FALSE;
   STAT0.STAT6 := FALSE;
   STAT0.STAT7 := FALSE;
   STAT0.STAT8 := FALSE;
   STAT0.STAT9 := FALSE;
   STAT0.STAT10 := TRUE;
   STAT0.STAT11 := FALSE;
   STAT0.STAT12 := FALSE;
   STAT0.STAT13 := FALSE;
   STAT0.STAT14 := FALSE;
   STAT0.STAT15 := FALSE;
   STAT0.STAT16 := FALSE;
   STAT0.STAT17[0] := W#16#0;
   STAT0.STAT17[1] := W#16#0;
   STAT0.STAT17[2] := W#16#0;
   STAT0.STAT17[3] := W#16#0;
   STAT0.STAT17[4] := W#16#0;
   STAT0.STAT17[5] := W#16#0;
   STAT0.STAT17[6] := W#16#0;
   STAT0.STAT17[7] := W#16#0;
   STAT18.STAT19 := 4296;
   STAT18.STAT20 := 3554;
   STAT18.STAT21 := 16961;
   STAT18.STAT22 := 17991;
   STAT18.STAT23 := -2580;
   STAT18.STAT24 := -1401;
   STAT18.STAT25 := -3129;
   STAT18.STAT26 := -2572;
   STAT18.STAT27 := 0;
   STAT18.STAT28 := 0;
   STAT29.STAT30 := -3944;
   STAT29.STAT31 := 11794;
   STAT29.STAT32 := -5083;
   STAT29.STAT33 := -5552;
   STAT29.STAT34 := -4763;
   STAT29.STAT35 := -5374;
   STAT29.STAT36 := 23843;
   STAT29.STAT37 := 24319;
   STAT29.STAT38 := 0;
   STAT29.STAT39 := 0;
   STAT40.STAT41 := 512;
   STAT40.STAT42 := 7338;
   STAT40.STAT43 := -442;
   STAT40.STAT44 := -671;
   STAT40.STAT45 := -1799;
   STAT40.STAT46 := -1968;
   STAT40.STAT47 := 18913;
   STAT40.STAT48 := 19376;
   STAT40.STAT49 := 0;
   STAT40.STAT50 := 0;
   STAT51.STAT52 := -17609;
   STAT51.STAT53 := 25459;
   STAT51.STAT54 := 2769;
   STAT51.STAT55 := 3114;
   STAT51.STAT56 := 3710;
   STAT51.STAT57 := 4098;
   STAT51.STAT58 := 25;
   STAT51.STAT59 := -586;
   STAT51.STAT60 := 0;
   STAT51.STAT61 := 0;
   STAT62.STAT63 := 0;
   STAT62.STAT64 := 0;
   STAT62.STAT65 := 0;
   STAT62.STAT66 := 0;
   STAT62.STAT67 := 0;
   STAT62.STAT68 := 0;
   STAT62.STAT69 := 0;
   STAT62.STAT70 := 0;
   STAT62.STAT71 := 0;
   STAT62.STAT72 := 0;
   STAT73.STAT74 := 0;
   STAT73.STAT75 := 0;
   STAT73.STAT76 := 0;
   STAT73.STAT77 := 0;
   STAT73.STAT78 := 0;
   STAT73.STAT79 := 0;
   STAT73.STAT80 := 0;
   STAT73.STAT81 := 0;
   STAT73.STAT82 := 0;
   STAT73.STAT83 := 0;
   STAT84.STAT85 := 0;
   STAT84.STAT86 := 0;
   STAT84.STAT87 := 0;
   STAT84.STAT88 := 0;
   STAT84.STAT89 := 0;
   STAT84.STAT90 := 0;
   STAT84.STAT91 := 0;
   STAT84.STAT92 := 0;
   STAT84.STAT93 := 0;
   STAT84.STAT94 := 0;
END_DATA_BLOCK

DATA_BLOCK DB 150
VERSION : 0.1


  STRUCT
   STAT0 : DWORD ;
   STAT1 : DWORD ;
   STAT2 : REAL ;
   STAT3 : REAL ;
   STAT4 : REAL ;
   STAT5 : WORD ;
   STAT6 : WORD ;
   STAT7 : WORD ;
   STAT8 : WORD ;
   STAT9 : DWORD ;
   STAT10 : REAL ;
   STAT11 : REAL ;
   STAT12 : REAL ;
   STAT13 : WORD ;
   STAT14 : WORD ;
   STAT15 : WORD ;
   STAT16 : WORD ;
   STAT17 : DWORD ;
   STAT18 : REAL ;
   STAT19 : REAL ;
   STAT20 : REAL ;
   STAT21 : WORD ;
   STAT22 : WORD ;
   STAT23 : WORD ;
   STAT24 : WORD ;
   STAT25 : DWORD ;
   STAT26 : REAL ;
   STAT27 : REAL ;
   STAT28 : REAL ;
   STAT29 : WORD ;
   STAT30 : WORD ;
   STAT31 : WORD ;
   STAT32 : WORD ;
   STAT33 : DWORD ;
   STAT34 : REAL ;
   STAT35 : REAL ;
   STAT36 : REAL ;
   STAT37 : WORD ;
   STAT38 : WORD ;
   STAT39 : WORD ;
   STAT40 : WORD ;
   STAT41 : DWORD ;
   STAT42 : REAL ;
   STAT43 : REAL ;
   STAT44 : REAL ;
   STAT45 : WORD ;
   STAT46 : WORD ;
   STAT47 : WORD ;
   STAT48 : WORD ;
   STAT49 : DWORD ;
   STAT50 : REAL ;
   STAT51 : REAL ;
   STAT52 : REAL ;
   STAT53 : WORD ;
   STAT54 : WORD ;
   STAT55 : WORD ;
   STAT56 : WORD ;
   STAT57 : DWORD ;
   STAT58 : REAL ;
   STAT59 : REAL ;
   STAT60 : REAL ;
   STAT61 : WORD ;
   STAT62 : WORD ;
   STAT63 : WORD ;
   STAT64 : WORD ;
   STAT65 : DWORD ;
   STAT66 : REAL ;
   STAT67 : REAL ;
   STAT68 : REAL ;
   STAT69 : WORD ;
   STAT70 : WORD ;
   STAT71 : WORD ;
   STAT72 : WORD ;
   STAT73 : DWORD ;
   STAT74 : REAL ;
   STAT75 : REAL ;
   STAT76 : REAL ;
   STAT77 : WORD ;
   STAT78 : WORD ;
   STAT79 : WORD ;
   STAT80 : WORD ;
   STAT81 : DWORD ;
   STAT82 : WORD ;
   STAT83 : WORD ;
   STAT84 : WORD ;
   STAT85 : WORD ;
   STAT86 : WORD ;
   STAT87 : WORD ;
   STAT88 : WORD ;
   STAT89 : WORD ;
   STAT90 : WORD ;
   STAT91 : WORD ;
   STAT92 : WORD ;
   STAT93 : WORD ;
   STAT94 : WORD ;
   STAT95 : WORD ;
   STAT96 : WORD ;
   STAT97 : BYTE ;
   STAT98 : BYTE ;
   STAT99 : BYTE ;
   STAT100 : BYTE ;
   STAT101 : BOOL ;
   STAT102 : BYTE ;
   STAT103 : BYTE ;
   STAT104 : BYTE ;
   STAT105 : WORD ;
   STAT106 : DINT ;
   STAT107 : DINT ;
   STAT108 : DINT ;
   STAT109 : REAL ;
   STAT110 : REAL ;
   STAT111 : REAL ;
   STAT112 : REAL ;
   STAT113 : REAL ;
   STAT114 : REAL ;
   STAT115 : REAL ;
   STAT116 : REAL ;
   STAT117 : REAL ;
   STAT118 : REAL ;
   STAT119 : REAL ;
   STAT120 : REAL ;
   STAT121 : REAL ;
   STAT122 : REAL ;
   STAT123 : REAL ;
   STAT124 : REAL ;
   STAT125 : REAL ;
   STAT126 : REAL ;
   STAT127 : REAL ;
   STAT128 : REAL ;
   STAT129 : REAL ;
   STAT130 : REAL ;
  END_STRUCT ;
BEGIN
   STAT0 := DW#16#800;
   STAT1 := DW#16#0;
   STAT2 := 2.054582e+003;
   STAT3 := -5.394847e+003;
   STAT4 := -1.542431e+003;
   STAT5 := W#16#0;
   STAT6 := W#16#0;
   STAT7 := W#16#0;
   STAT8 := W#16#0;
   STAT9 := DW#16#2;
   STAT10 := 2.149658e-001;
   STAT11 := 8.890132e+002;
   STAT12 := -1.498335e+003;
   STAT13 := W#16#0;
   STAT14 := W#16#0;
   STAT15 := W#16#0;
   STAT16 := W#16#0;
   STAT17 := DW#16#200;
   STAT18 := 9.505859e+000;
   STAT19 := 8.919878e+002;
   STAT20 := -1.090076e+003;
   STAT21 := W#16#0;
   STAT22 := W#16#0;
   STAT23 := W#16#0;
   STAT24 := W#16#0;
   STAT25 := DW#16#200;
   STAT26 := -1.638507e+003;
   STAT27 := 8.918486e+002;
   STAT28 := -2.388569e+003;
   STAT29 := W#16#0;
   STAT30 := W#16#0;
   STAT31 := W#16#0;
   STAT32 := W#16#0;
   STAT33 := DW#16#200;
   STAT34 := 0.000000e+000;
   STAT35 := 0.000000e+000;
   STAT36 := 0.000000e+000;
   STAT37 := W#16#0;
   STAT38 := W#16#0;
   STAT39 := W#16#0;
   STAT40 := W#16#0;
   STAT41 := DW#16#0;
   STAT42 := 0.000000e+000;
   STAT43 := 0.000000e+000;
   STAT44 := 0.000000e+000;
   STAT45 := W#16#0;
   STAT46 := W#16#0;
   STAT47 := W#16#0;
   STAT48 := W#16#0;
   STAT49 := DW#16#0;
   STAT50 := 0.000000e+000;
   STAT51 := 0.000000e+000;
   STAT52 := 0.000000e+000;
   STAT53 := W#16#0;
   STAT54 := W#16#0;
   STAT55 := W#16#0;
   STAT56 := W#16#0;
   STAT57 := DW#16#0;
   STAT58 := 0.000000e+000;
   STAT59 := 0.000000e+000;
   STAT60 := 0.000000e+000;
   STAT61 := W#16#0;
   STAT62 := W#16#0;
   STAT63 := W#16#0;
   STAT64 := W#16#0;
   STAT65 := DW#16#0;
   STAT66 := 0.000000e+000;
   STAT67 := 0.000000e+000;
   STAT68 := 0.000000e+000;
   STAT69 := W#16#0;
   STAT70 := W#16#0;
   STAT71 := W#16#0;
   STAT72 := W#16#0;
   STAT73 := DW#16#0;
   STAT74 := 0.000000e+000;
   STAT75 := 0.000000e+000;
   STAT76 := 0.000000e+000;
   STAT77 := W#16#0;
   STAT78 := W#16#0;
   STAT79 := W#16#0;
   STAT80 := W#16#0;
   STAT81 := DW#16#0;
   STAT82 := W#16#3;
   STAT83 := W#16#33;
   STAT84 := W#16#0;
   STAT85 := W#16#3;
   STAT86 := W#16#2DE;
   STAT87 := W#16#0;
   STAT88 := W#16#3;
   STAT89 := W#16#763;
   STAT90 := W#16#792;
   STAT91 := W#16#3;
   STAT92 := W#16#B4;
   STAT93 := W#16#C5;
   STAT94 := W#16#3;
   STAT95 := W#16#FFD4;
   STAT96 := W#16#FFBD;
   STAT97 := B#16#0;
   STAT98 := B#16#FF;
   STAT99 := B#16#0;
   STAT100 := B#16#14;
   STAT101 := FALSE;
   STAT102 := B#16#0;
   STAT103 := B#16#0;
   STAT104 := B#16#FF;
   STAT105 := W#16#0;
   STAT106 := L#1770;
   STAT107 := L#884;
   STAT108 := L#1006;
   STAT109 := 8.200000e+001;
   STAT110 := 8.100000e+001;
   STAT111 := 2.490000e+002;
   STAT112 := 1.130000e+003;
   STAT113 := -3.130000e+002;
   STAT114 := 3.330000e+002;
   STAT115 := 1.183000e+003;
   STAT116 := -3.430000e+002;
   STAT117 := 3.600000e+002;
   STAT118 := 1.505000e+003;
   STAT119 := 7.200000e+002;
   STAT120 := 1.200000e+003;
   STAT121 := 2.156000e+003;
   STAT122 := 1.283000e+003;
   STAT123 := -1.842000e+003;
   STAT124 := -2.346744e+000;
   STAT125 := 2.176595e-001;
   STAT126 := 1.453762e+001;
   STAT127 := 0.000000e+000;
   STAT128 := 0.000000e+000;
   STAT129 := 0.000000e+000;
   STAT130 := 0.000000e+000;
END_DATA_BLOCK

DATA_BLOCK DB 200
VERSION : 0.1


  STRUCT
   STAT0 : DATE_AND_TIME  := DT#95-1-1-0:0:0.000;
   STAT1 : DATE_AND_TIME  := DT#95-1-1-0:0:0.000;
   STAT2 : INT ;
   STAT3 : DATE  := D#1995-1-1;
   STAT4 : TIME_OF_DAY ;
   STAT5 : INT ;
   STAT6 : BYTE ;
  END_STRUCT ;
BEGIN
   STAT0 := DT#95-1-1-0:0:0.000;
   STAT1 := DT#01-5-4-23:48:57.905;
   STAT2 := 0;
   STAT3 := D#1995-1-1;
   STAT4 := TOD#0:0:0.000;
   STAT5 := 0;
   STAT6 := B#16#0;
END_DATA_BLOCK

FUNCTION_BLOCK FB 250
VERSION : 1.1


